      def clipWhenLowerLimitIsLessThanHigher(outputScaledValue, outputRange):
          if (outputScaledValue < outputRange[0]):
              return outputRange[0]
          elif (outputScaledValue > outputRange[1]):
              return outputRange[1]
          else:
              return outputScaledValue
          end
      end

      slope = computeSlope(rawRange, scaledRange)
      intercept = computeIntercept(slope, rawRange, scaledRange)
      scaledValue = slope * value + intercept
      return clipScaledValue(scaledValue, scaledRange)
  end

  def limit(value, range):
      return scale(value, range, range)
  end


  rq_init_comm_if_connected(9, "1")
  rq_init_comm_if_connected(2, "2")
  rq_init_comm_if_connected(3, "3")
  rq_init_comm_if_connected(4, "4")
  rq_print_connected_grippers()
  rq_gripper_communication_thread = run rq_gripper_communication()
  set_closed_norm(97.6470588235294, 1)
  set_open_norm(1.1764705882352942, 1)
  set_closed_mm(0.0, 1)
  set_open_mm(53.0, 1)
  set_closed_norm(100.0, 2)
  set_open_norm(0.0, 2)
  set_closed_mm(0.0, 2)
  set_open_mm(50.0, 2)
  set_closed_norm(100.0, 3)
  set_open_norm(0.0, 3)
  set_closed_mm(0.0, 3)
  set_open_mm(50.0, 3)
  set_closed_norm(100.0, 4)
  set_open_norm(0.0, 4)
  set_closed_mm(0.0, 4)
  set_open_mm(50.0, 4)
  rq_current_limit_enabled = False
  while(not rq_gripper_communication_thread_started):
      sync()
  end
  # end: URCap Installation Node
  # begin: URCap Installation Node
  #   Source: OPC UA, 2.0.2, Rocketfarm AS
  #   Type: OPC UA
  global opcua_daemon = rpc_factory("xmlrpc", "http://127.0.0.1:40409/RPC2")
  def opcua_client_connect(address):
  return opcua_daemon.client_connect(address)
  end
  def opcua_client_get_id(client_name):
  return opcua_daemon.client_get_id(client_name)
  end
  def opcua_client_try_connect(client_id):
  opcua_result = False
  if (opcua_daemon.client_connect(client_id)):
  sleep(0.01)
  opcua_result = opcua_daemon.client_is_connected(client_id)
  opcua_retry = 10
  while ( (not opcua_result) and (opcua_retry > 0) ):
  sleep(0.1)
  opcua_result = opcua_daemon.client_is_connected(client_id)
  opcua_retry = opcua_retry - 1
  end
  end
  return opcua_result
  end
  def opcua_client_disconnect(client_id):
  return opcua_daemon.client_disconnect(client_id)
  end
  def opcua_client_is_connected(client_id):
  return opcua_daemon.client_is_connected(client_id)
  end
  def opcua_client_read_byid(client_id, namespace_id, variable_id):
  return opcua_daemon.client_read_variable_by_id(client_id, namespace_id, variable_id)
  end
  def opcua_client_read_byname(client_id, namespace_id, variable_name):
  return opcua_daemon.client_read_variable_by_name(client_id, namespace_id, variable_name)
  end
  def opcua_client_write_byid(client_id, namespace_id, variable_id, variable_value):
  return opcua_daemon.client_write_variable_by_id(client_id, namespace_id, variable_id, variable_value)
  end
  def opcua_client_write_byname(client_id, namespace_id, variable_name, variable_value):
  return opcua_daemon.client_write_variable_by_name(client_id, namespace_id, variable_name, variable_value)
  end
  def opcua_client_last_error(client_id):
  return opcua_daemon.client_get_last_error(client_id)
  end
  def opcua_server_read_byname(variable_name):
  return opcua_daemon.server_read_variable_by_name(variable_name)
  end
  def opcua_server_write_byname(variable_name, variable_value):
  return opcua_daemon.server_write_variable_by_name(variable_name, variable_value)
  end
  def opcua_server_last_error():
  return opcua_daemon.server_get_last_error()
  end
  def opcua_error_to_string(errorCode):
  return opcua_daemon.error_code_to_string(errorCode)
  end
  # end: URCap Installation Node
  global CAM_Pose=p[0,0,0,0,0,0]
  global CAM_Relation=""
  global CMD_Abort=  False
  global CMD_Clear=  False
  global CMD_Reset=  False
  global CMD_Start=  False
  global CMD_Suspend=  False
  global CMD_Unhold=  False
  global CMD_Unsuspend=  False
  global CNT_Rack_Output=0
  global FNC_Freedrive=  False
  global PRC_TubCounter=0
  global STP=0
  global easyPickCount=0
  global easyPickCount_4=0
  global easyPickCount_6=0
  global easyPickCount_7=0
  global easyPickNoObj=0
  global easyPickNoObj_4=0
  global easyPickNoObj_6=0
  global easyPickNoObj_7=0
  global easyPickParts=0
  global easyPickParts_4=0
  global easyPickParts_6=0
  global easyPickParts_7=0
  global Container_mid_1_p=p[-.379239199143, -.127191311915, .299999999998, .000000000046, -.000000000021, -1.247199999994]
  global Container_mid_1_q=[-2.477408934449926, -1.2969853503591224, -1.875639182904262, -1.539621866126728, 1.5731943360401213, -2.8009955944022717]
  global Container_capt_p=p[-.525590029047, .407247642794, .411588185841, -.000000000107, .000000000065, -2.896148821900]
  global Container_capt_q=[-3.5968351615224767, -2.0050156108707204, -0.8176271154495112, -1.8895759482008394, 1.5730967555598792, -2.2743681102957645]
  global Waypoint_51_p=p[-.335468094724, -.217855817953, .299999999998, .000000000047, -.000000000014, -.994837065669]
  global Waypoint_51_q=[-2.2250460001249586, -1.2969853503591224, -1.875639182904262, -1.539621866126728, 1.573194336040121, -2.800995594402271]
  global Waypoint_13_p=p[-.479450777041, .284140798427, .125270103493, -.276792173670, 2.098433187455, -2.121256516887]
  global Waypoint_13_q=[-2.8915050665484827, -1.9549266300597132, -2.2318272590637207, -1.6654960117735804, 0.020810842514038086, -0.4019392172442835]
  global Waypoint_70_p=p[-.472820924464, .292439826304, .207418370234, -.259787347864, -2.053484648504, 2.070709755662]
  global Waypoint_70_q=[-2.969927421603815, -2.07168115810532, -1.6835546062719366, -2.4953958198513964, 0.4489790927922641, -0.005578998612037367]
  global Waypoint_2_p=p[-.312961047461, -.152991312519, .223609826854, -.745314530454, -1.713873240489, 1.673341715282]
  global Waypoint_2_q=[-2.3560472170459192, -2.183784624139303, -1.4583134651184082, -2.6435262165465296, 1.6522362232208252, 0.043451953679323196]
  global Waypoint_3_p=p[-.113749865836, -.390110151572, .317307487562, -.519383711706, -.839884211339, 1.756868173041]
  global Waypoint_3_q=[-1.8909733931170862, -1.720626016656393, -1.5115610361099243, -2.1240560017027796, 2.1809096336364746, 0.7227501273155212]
  global Waypoint_15_p=p[.029144035010, -.436802470887, .327885032028, -.521560953301, -.623641814548, 1.862659450154]
  global Waypoint_15_q=[-1.564817253743307, -1.556895188321807, -1.6826975345611572, -1.6944714985289515, 2.2362685203552246, 1.117417335510254]
  global Waypoint_14_p=p[.068712235638, -.569419545175, .285215357659, -.679242949116, -.712065334485, 1.394044574094]
  global Waypoint_14_q=[-1.5731792953485346, -1.8029235103747094, -1.6781008808776736, -1.2218450646111982, 2.4719572998240125, 1.6394218026856375]
  global Waypoint_4_p=p[-.047220457210, -.557624911767, .136370962514, -.679242949107, -.712065334475, 1.394044574096]
  global Waypoint_4_q=[-1.7740079055958748, -2.0023561428872334, -1.7577251142892676, -1.18903287716154, 2.4487287370345143, 1.322902469273079]
  global Waypoint_25_p=p[.065436479647, -.569388431626, .287820755049, -.679242949185, -.712065334557, 1.394044574070]
  global Waypoint_25_q=[-1.5789263550890595, -1.8020194754825436, -1.6702557537748035, -1.237882536889547, 2.471995808083492, 1.6301087487321393]
  global Waypoint_39_p=p[.137772150180, -.577759956854, .299999999946, .000000000217, -.000000000207, -1.594351842625]
  global Waypoint_39_q=[-1.108978697428574, -1.776486680444405, -1.413737665315093, -1.5218908901738937, 1.5733062372356947, -1.0863866394180182]
  global Waypoint_41_p=p[.074222967010, -.565641640647, .234620140366, -.516884386806, .529223682286, -1.529619060506]
  global Waypoint_41_q=[-0.9596722604286052, -1.8767069964135548, -1.4892746174057256, -1.7813862040292285, 1.0520698599867686, -0.8199687448260349]
  global Waypoint_40_p=p[.039987741677, -.564832865048, .191055405868, -.767560686167, .343136533060, -2.241315728308]
  global Waypoint_40_q=[-1.0070649180116558, -1.8745927522477324, -1.6139175023195245, -1.6337474788493545, 1.032708081143138, -0.11587278312988403]
  global Waypoint_42_p=p[.041363380882, -.564865360786, .192805844739, .278500165520, .624117100927, .762272396553]
  global Waypoint_42_q=[-1.0050718976263102, -1.8744386685524779, -1.609151451954446, -1.6399653140247947, 1.0334006002355505, -3.254032861659603]
  global Waypoint_43_p=p[.041363380886, -.564865360780, .192805844755, .854271020883, .226833028600, 2.453002871494]
  global Waypoint_43_q=[-1.0050567614299233, -1.874341297657562, -1.6092945416026048, -1.6397580431809713, 1.0333661149462194, -5.0371728933995605]
  global Waypoint_44_p=p[.040882892233, -.564854254876, .192193763716, .110913882012, .659173708659, .275719738520]
  global Waypoint_44_q=[-1.0057704811530535, -1.8745207681598055, -1.6107765025572558, -1.637858394640876, 1.033164860873599, -2.7487836132940755]
  global Waypoint_45_p=p[.042647731639, -.564895808997, .194439423694, -.451694728506, .563172064821, -1.343350300184]
  global Waypoint_45_q=[-1.0032860829914387, -1.8741561795270565, -1.6048483308761785, -1.6453689714776623, 1.0342050634514657, -1.06078829880322]
  global Waypoint_46_p=p[.099944144487, -.566244126804, .267342790130, -.451694834765, .563172023386, -1.343350532536]
  global Waypoint_46_q=[-0.9257438092434924, -1.889970530402497, -1.3828165217629076, -1.8916791100652528, 1.0664350961373816, -0.9805910833329659]
  global Waypoint_47_p=p[.099944144444, -.566244126727, .267342790273, -.101742139519, .058679218003, -1.457888523314]
  global Waypoint_47_q=[-1.1112623176383014, -1.729989471869196, -1.5530029871033957, -1.4442770617454777, 1.4670579052775654, -1.2224020460061675]
  global Waypoint_48_p=p[-.136182767566, -.647487115908, .294247768372, -.101742139549, .058679218020, -1.457888523312]
  global Waypoint_48_q=[-1.532196177857717, -1.9115932455375173, -1.2651848069729779, -1.5055651746702665, 1.4703193777418382, -1.646379689188814]
  global Waypoint_49_p=p[-.159024328559, -.641021381179, .047691706070, -.000000000033, -.000000000027, -1.457897102937]
  global Waypoint_49_q=[-1.6098490079965062, -2.1164987141784586, -1.6156631902166785, -0.9800092198841526, 1.573231151532669, -1.722204302767242]
  global Waypoint_50_p=p[-.159024328558, -.641021381151, .291114489351, -.000000000033, -.000000000027, -1.457897102937]
  global Waypoint_50_q=[-1.609190265995684, -1.9426985888940234, -1.2189094859258596, -1.55056435122874, 1.5734384912955113, -1.7235116759964022]
  global Waypoint_53_p=p[-.050111345339, -.357608435610, .335880801283, .034180375734, .020280946727, -.284888945062]
  global Waypoint_53_q=[-1.3262308189700454, -1.2221767968893875, -1.8246061249803773, -1.7046285947349489, 1.567288986353525, -2.612420684434543]
  global Spatula_above_p=p[.241880327671, -.243077591927, .290283157642, .000026293989, -.000477463062, 3.067686800856]
  global Spatula_above_q=[-0.3881264518731289, -1.1433094134493045, -1.996913957798169, -1.572030383936684, 1.5734346414190374, 1.2567789862982233]
  global Spatula_pick_p=p[.240292635430, -.243077591534, .189212061148, .000026293987, -.000477463065, 3.067686800855]
  global Spatula_pick_q=[-0.39083408330539005, -1.1777602778656497, -2.2383115866577645, -1.2961817529600745, 1.573403050820434, 1.2551372216266965]
  global container_start_p=p[.200650292946, -.570238751958, .366326773614, 1.360500828661, .021700128770, 2.681649891414]
  global container_start_q=[-0.7669977765142582, -2.188996679669204, -0.7412727239230232, -2.581362891432544, 1.0193601740278728, 1.1884911920528847]
  global container_wp_1_p=p[.170613637794, -.572150573676, .294509026043, 1.259497117139, -.008270589399, 2.787717865625]
  global container_wp_1_q=[-0.8129253370121727, -2.0726598902108755, -1.0846040680899218, -2.2403146195823957, 1.0281191187839607, 1.0435744211830564]
  global Waypoint_55_p=p[.077280900603, -.567308602990, .212067617714, 1.259497117148, -.008270589399, 2.787717865619]
  global Waypoint_55_q=[-0.9181858327853867, -1.9744793804952083, -1.4540279077890048, -1.9155621911627945, 0.9643238328181578, 0.9457250675800015]
  global Waypoint_56_p=p[.135568164031, -.570867938153, .245215470413, 1.476861317558, -.018269607491, 2.679642659499]
  global Waypoint_56_q=[-0.8259784040282607, -2.108036981522602, -1.2111990877342924, -2.2405969375728745, 0.9451797152137279, 1.125710531287379]
  global Waypoint_74_p=p[.164827890887, -.574638012411, .193751361296, 2.053636896063, -.046507887560, 2.274278266449]
  global Waypoint_74_q=[-0.7657213433975762, -2.450387120010788, -0.9886183070290357, -2.7078095590939375, 0.8831550681477878, 1.5106229631053527]
  global ftr_scoop2_p=p[.194287054614, -.495779761333, .282072128495, -.179029871953, 1.612108092436, -.016025695011]
  global ftr_scoop2_q=[-0.5957383150173561, -2.264100500923713, -1.1936887184643812, -2.8893702964346097, 0.8750688478879766, -1.4109843517598684]
  global aftr_scoo3_p=p[-.289759911340, -.315385007342, .303743796282, .159961590809, 1.627415489603, -.344855744095]
  global aftr_scoo3_q=[-1.3374747909924949, -1.6809733407851706, -1.9857606509106667, -2.713564895186775, 0.5589807453366573, -1.3631067603374376]
  global Waypoint_60_p=p[-.013316432876, -.544772031582, .383371643081, 2.208233379808, .037543335712, 2.097559881761]
  global Waypoint_60_q=[-0.9328326161883087, -2.0999933666355775, -1.1958015693111372, -3.060905141293654, 0.690378518537611, 1.7121940951337198]
  global Waypoint_61_p=p[-.412188693372, -.356446875193, .383371643081, 1.751740964455, -.739956256289, 1.600691174920]
  global Waypoint_61_q=[-1.766185342973321, -2.0999933666355775, -1.1958015693111372, -3.060905141293654, 0.690378518537611, 1.7121940951337198]
  global Waypoint_75_p=p[-.343126484123, -.342779621892, .335357223804, .359429517288, 1.600352990741, -.365083732359]
  global Waypoint_75_q=[-1.517806275013295, -1.8136828056045395, -1.737638081810795, -2.8432599585466436, 0.5149430839716123, -1.4579122147201877]
  global aftr_scoop1_p=p[.138503854266, -.514479969882, .214153672011, -.134825326227, 1.559916297527, -.059196589314]
  global aftr_scoop1_q=[-0.6880464314785328, -2.2689986529709643, -1.3310176475983653, -2.673087158390708, 0.8340516295138949, -1.4557846480003231]
  global After_disp_3_p=p[.125934854156, -.585611107804, .299545938076, .959554236104, -.134386766509, 2.880651774211]
  global After_disp_3_q=[-0.9434480594885066, -2.016473586333989, -1.1036579072158617, -2.096459283015281, 1.1479556364931514, 0.8433331387406042]
  global Waypoint_62_p=p[-.542658707241, -.114281911009, .251261544113, 1.813043609523, -.679411528034, 1.655271622964]
  global Waypoint_62_q=[-2.158300033470912, -1.9418836862428677, -1.8142999147147894, -2.778920736683023, 0.21900622104017292, 1.8983390235012934]
  global Waypoint_63_p=p[.101294795191, -.465376052375, .381756220355, .972633305146, -.158447626639, 2.887199602585]
  global Waypoint_63_q=[-0.8528172446194038, -1.7393709485118478, -1.2544079521837954, -2.2703112963960628, 1.1965892397133469, 0.91867216443391]
  global Start_p=p[-.033064633790, -.365398531763, .389873206922, .000000000001, .000000000001, 2.725785203584]
  global Start_q=[-1.287596562866887, -1.232866726886848, -1.6880113260231102, -1.7912103151657988, 1.5729028131945846, 0.6981423183093938]
  global Waypoint_76_p=p[-.479450777041, .284140798427, .125270103493, -.276792173670, 2.098433187454, -2.121256516887]
  global Waypoint_76_q=[-2.891505066548503, -1.9549266300590151, -2.231827259067863, -1.6654960117542226, 0.020810842514162875, -0.4019392172601952]
  global PowderA_wayp1_p=p[-.472820924474, .292439826233, .207418370237, -.137787250486, 2.177332259632, -2.152029714756]
  global PowderA_wayp1_q=[-2.911134078210732, -1.90240864358569, -1.968768330510411, -2.500365101593811, 0.11427687110891149, 0.0958980389250167]
  global Waypoint_80_p=p[-.303921889165, -.326082520111, .297721580072, -.584846481381, 1.914382606328, -1.960922301253]
  global Waypoint_80_q=[-1.6364180099980672, -2.041258366871811, -1.472153549517767, -2.7572808013122696, 0.9684003593854582, 0.047163023020230455]
  global Decapp_above_p=p[-.013480295948, -.359153355979, .266194408367, -.879653555922, 1.646336924805, -1.709111068605]
  global Decapp_above_q=[-0.9632157249872035, -2.0163405763031657, -1.5968194594157152, -2.6579215719847085, 1.251243398585566, 0.047906446502667066]
  global Decapp_place_p=p[-.013480295848, -.359153356116, .158558645017, -.879653554904, 1.646336919751, -1.709111066446]
  global Decapp_place_q=[-0.9633419174801583, -2.157735564881908, -1.695182597572722, -2.418253553201909, 1.2517436353048952, 0.04819090596102882]
  global Waypoint_78_p=p[-.051450028091, -.519555688329, .365718563414, -1.287302938145, 1.077637394477, -1.218524965834]
  global Waypoint_78_q=[-0.9214276262416012, -1.8899696965062578, -1.4939326452510562, -2.840015661555725, 0.5585157189668353, 0.033997638875617575]
  global Waypoint_81_p=p[-.030847790230, -.346237542439, .241203613248, .000000000000, .000000000000, .000000000000]
  global Waypoint_81_q=[-1.265848516232941, -1.1652881302267932, -2.11003646605462, -1.4369228603041853, 1.573284436504383, -2.835929896730388]
  global Waypoint_79_p=p[-.030847972829, -.346235312674, .229874122470, .000000000000, .000000000000, .000000000000]
  global Waypoint_79_q=[-1.2659333103898618, -1.1699230683425625, -2.1365870669440055, -1.4057372655396474, 1.5732787836040316, -2.8358953794066757]
  global Waypoint_82_p=p[-.031079593487, -.346547394534, .293012696855, -.000011575267, -.000017731224, -.000713984074]
  global Waypoint_82_q=[-1.2664169521879751, -1.1572597700415788, -1.982185304253158, -1.5727862504184884, 1.5732673022058234, -2.83632822711502]
  global Cap_above_p=p[-.163602500478, -.618357694237, .258271116068, .000026793591, -.000032305852, -.969382601663]
  global Cap_above_q=[-1.6181634639269902, -1.896432778341337, -1.3662765317923142, -1.449515114018281, 1.5734416863575176, -2.220489512402157]
  global Cap_Place_p=p[-.153420247224, -.637174247221, .035295616791, .000000000002, -.000000000002, -1.457849918374]
  global Cap_Place_q=[-1.6014084627078784, -2.123124488207292, -1.6429187572395012, -0.946127085055064, 1.573175527437006, -1.7136981844648291]
  global OP_PowderA2_p=p[.009371277507, -.409434369247, .294169017766, -.823281033205, 1.709410851243, -1.698303593897]
  global OP_PowderA2_q=[-0.9994544761745754, -2.1395254572673217, -1.3437567783153916, -2.8143375616690456, 1.2617899549595724, 0.019614613715634555]
  global OP_PowderA_abov_p=p[-.012145216791, -.363335041455, .315325728178, -.777135478411, 1.752984823781, -1.740925591659]
  global OP_PowderA_abov_q=[-1.01634425044037, -2.024785947780374, -1.4658894155189923, -2.8070189735738786, 1.3091674480404514, 0.020022086766872782]
  global OP_PowderA_pick_p=p[-.012145216707, -.363335041590, .179898787547, -.777135478413, 1.752984823781, -1.740925591659]
  global OP_PowderA_pick_q=[-1.0165129229305911, -2.176980100858497, -1.6127054339661555, -2.5080740815244567, 1.3098787614888208, 0.020270375244195882]
  global Op_PowA_wP_p=p[-.173727579245, -.372934016396, .295116627479, -.972390492433, 1.540962074418, -1.548745344994]
  global Op_PowA_wP_q=[-1.1740587397768483, -1.865656321049359, -1.7426943793777419, -2.679427276872525, 0.8588908769087338, 0.017944699631825187]
  global Waypoint_1_p=p[-.451048883256, -.340589460864, .308223661552, .097058877504, .091048998701, -1.578386010942]
  global Waypoint_1_q=[-2.222400490437643, -1.7554131946959437, -1.398173213005066, -1.6564461193480433, 1.5042352676391602, -2.2106884161578577]
  global Spatula_otw_p=p[-.038472058237, -.263141484147, .425351216717, -.000441582511, -.000128175490, 3.034387645854]
  global Spatula_otw_q=[-1.1888947506684495, -1.0083288774886814, -1.7052227056065874, -1.9984805067363443, 1.5730180972985317, 0.48793409320312264]
  global pick_spat_L_abv_p=p[.247376339171, -.151300871293, .298405979617, .000026293989, -.000477463062, 3.067686800856]
  global pick_spat_L_abv_q=[-0.07082187843937948, -0.9918336120099029, -2.048431407771396, -1.6719226065707566, 1.5735148227092874, 1.5739821706892307]
  global spat_L_pick_p=p[.244425006707, -.151048053384, .192288246285, .000026293989, -.000477463065, 3.067686800855]
  global spat_L_pick_q=[-0.07170850917614935, -0.9939169317558161, -2.3190151588645502, -1.3992549297298966, 1.573619586467819, 1.5742112847515592]
  global spat_L_lift_p=p[.247500241215, -.151291104039, .242146826477, .000026293989, -.000477463064, 3.067686800855]
  global spat_L_lift_q=[-0.07132168213116863, -0.9873531406871798, -2.1938095635783172, -1.531024644535787, 1.5736129628476565, 1.5740661231239859]
  global spat_L_side_p=p[.251772314117, -.093610100391, .242165935204, .000026293989, -.000477463064, 3.067686800855]
  global spat_L_side_q=[0.16311920731341095, -0.9159674867544636, -2.2202625845173465, -1.5759061264106862, 1.5736725172206427, 1.8084579794657634]
  global spat_L_up_p=p[.248631729748, -.094370561652, .425351216716, .000026293989, -.000477463065, 3.067686800855]
  global spat_L_up_q=[0.16435650344985986, -1.008385469590376, -1.7051729211515223, -1.9985780211252369, 1.5729805495343943, 1.8078858605162342]
  global spat_M_up_p=p[.246651483123, -.200758466677, .427983242435, .000026293988, -.000477463066, 3.067686800854]
  global spat_M_up_q=[-0.2488061154947081, -1.1388154682286178, -1.6405006043284098, -1.932909670500866, 1.5729930693357987, 1.394694958078517]
  global spat_M_pick_p=p[.243754824031, -.195909855689, .192274495860, .000026293989, -.000477463063, 3.067686800855]
  global spat_M_pick_q=[-0.2371047546337337, -1.0815273547611497, -2.2806002623741977, -1.3500947192370933, 1.573515135501001, 1.4088438823663394]
  global spat_S_up_p=p[.250500617207, -.246905508589, .391583682111, .000026293987, -.000477463068, 3.067686800854]
  global spat_S_up_q=[-0.3880360419879594, -1.1962881911765244, -1.7058643812256875, -1.8101014540154097, 1.5731545967396166, 1.2558061200976702]
  global spat_S_pick_p=p[.245173607467, -.244249950907, .193022226997, .000026293988, -.000477463064, 3.067686800854]
  global spat_S_pick_q=[-0.38836215799357987, -1.1880037605751017, -2.222350098157584, -1.30189927792612, 1.5733998957551099, 1.2575641527417636]
  def Sub_Vision_V18():
    $ 714 "Sub_Vision_V18" "noBreak"
    $ 715 "PreSettings"
    $ 716 "CAM_LM_Detected≔ False "
    global CAM_LM_Detected=  False
    $ 717 "CAM_Captures≔0"
    global CAM_Captures=0
    $ 718 "CAM_Pose≔p[0,0,0,0,0,0]"
    global CAM_Pose=p[0,0,0,0,0,0]
    $ 719 "CAM_LM_Refinmnt≔ False "
    global CAM_LM_Refinmnt=  False
    $ 720 "CAM_LM_Refined≔ False "
    global CAM_LM_Refined=  False
    $ 721 "CAM_LM_Deviatn≔p[0,0,0,0,0,0]"
    global CAM_LM_Deviatn=p[0,0,0,0,0,0]
    $ 722 "CAM_LM_ID≔0"
    global CAM_LM_ID=0
    $ 723 "CAM_Done≔ False "
    global CAM_Done=  False
    $ 724 "CAM_CNT_Obj≔0"
    global CAM_CNT_Obj=0
    $ 725 "CAM_Result = []"
    CAM_Result = []
    $ 726 "OBJ_Detected≔ False "
    global OBJ_Detected=  False
    $ 727 "FRM_Reference≔p[0,0,0,0,0,0]"
    global FRM_Reference=p[0,0,0,0,0,0]
    $ 728 "'=========='"
    # '=========='
    $ 729 "Switch Action"
    switch_1 = Action
    $ 730 "Case 13"
    if (13 == switch_1):
    elif (15 == switch_1):
      $ 848 "Case 15"
    elif (131 == switch_1):
      $ 894 "Case 131"
      $ 895 "Read (SensoPart)"
      $ 896 "Action_Info≔'search for landmark'"
      global Action_Info="search for landmark"
      $ 897 "CAM_LM≔CAM_LMs[4]"
      global CAM_LM=CAM_LMs[4]
      $ 898 "CAM_Relation≔CAM_LM.capture_relation"
      global CAM_Relation=CAM_LM.capture_relation
      $ 899 "go to capture pose"
      $ 902 "If ITM_ID≟1 and JIG≟7"
      if (ITM_ID == 1  and  JIG == 7):
        $ 903 "PSE_T≔uLM_Cap_SSRack"
        global PSE_T=uLM_Cap_SSRack
      else:
        $ 904 "ElseIf ITM_ID≟5 and JIG≟7"
        if (ITM_ID == 5  and  JIG == 7):
          $ 905 "PSE_T≔FRM_Cap_SSRack"
          global PSE_T=FRM_Cap_SSRack
        else:
          $ 906 "ElseIf ITM_ID≟13 and JIG≟7"
          if (ITM_ID == 13  and  JIG == 7):
            $ 907 "PSE_T≔FRM_pick_rack_const"
            global PSE_T=p[-0.5568395192387274,0.34423986364170267,0.44698620470146266,-1.0069110132199915E-6,3.378712467497258E-5,-8.002029546773325E-6]
          else:
            $ 908 "ElseIf ITM_ID≟1 and JIG≟15"
            if (ITM_ID == 1 and JIG == 15):
              $ 909 "MoveJ"
              $ 910 "Container_mid_1" "breakAfter"
              movej(get_inverse_kin(Container_mid_1_p, qnear=Container_mid_1_q), a=1.3962634015954636, v=1.0471975511965976, r=0.05)
              $ 911 "Container_capt" "breakAfter"
              movej(get_inverse_kin(Container_capt_p, qnear=Container_capt_q), a=1.3962634015954636, v=1.0471975511965976)
              $ 912 "PSE_T≔FRM_Container_S_const"
              global PSE_T=p[-0.510412665574981,0.40064363362973565,0.41159789496794374,-1.1370875604168537E-5,-3.643547521609506E-6,-2.896122366208473]
            else:
              $ 913 "ElseIf ITM_ID≟1 and JIG≟16"
              if (ITM_ID == 1  and  JIG == 16):
                $ 914 "MoveJ"
                $ 915 "Waypoint_51" "breakAfter"
                movej(get_inverse_kin(Waypoint_51_p, qnear=Waypoint_51_q), a=1.3962634015954636, v=1.0471975511965976, r=0.05)
                $ 917 "PSE_T≔FRM_Weigh_scale_const"
                global PSE_T=p[-0.3454891122972868,0.06305469656946562,0.547028193804949,1.63274868305228E-4,-7.686242288056818E-5,-2.2741025165393225]
              else:
                $ 918 "ElseIf ITM_ID≟1 and JIG≟17"
                if (ITM_ID == 1  and  JIG == 17):
                  $ 919 "MoveJ"
                  $ 920 "Waypoint_51" "breakAfter"
                  movej(get_inverse_kin(Waypoint_51_p, qnear=Waypoint_51_q), a=1.3962634015954636, v=1.0471975511965976, r=0.05)
                  $ 922 "PSE_T≔FRM_Weigh_scale_const"
                  global PSE_T=p[-0.3454891122972868,0.06305469656946562,0.547028193804949,1.63274868305228E-4,-7.686242288056818E-5,-2.2741025165393225]
                else:
                  $ 923 "ElseIf ITM_ID≟1 and JIG≟21"
                  if (ITM_ID == 1  and  JIG == 21):
                    $ 924 "MoveJ"
                    $ 925 "Waypoint_51" "breakAfter"
                    movej(get_inverse_kin(Waypoint_51_p, qnear=Waypoint_51_q), a=1.3962634015954636, v=1.0471975511965976, r=0.05)
                    $ 927 "PSE_T≔FRM_PoTS_const"
                    global PSE_T=p[-0.5211683440725288,-0.17068665293155189,0.5469908617304544,2.009713344566374E-4,5.545167142016751E-6,-2.2342044673695503]
                  end
                end
              end
            end
          end
        end
      end
      $ 928 "do_transition(PSE_T, keep_rxry=False)"
      do_transition(PSE_T, keep_rxry=False)
      $ 929 "Set"
      set_tcp(p[0.0,0.0,0.161,3.1415,0.0,0.0])
      $ 930 "MoveJ"
      $ 931 "PSE_T" "breakAfter"
      movej(PSE_T, a=1.3962634015954636, v=1.7453292519943295)
      $ 932 "CAM_Pose≔get_actual_tcp_pose()"
      global CAM_Pose= get_actual_tcp_pose ()
      $ 933 "Loop  not CAM_Done and  not ERROR.FLAG and  not CMD_Stop"
      while (  not  CAM_Done  and    not  ERROR.FLAG  and    not  CMD_Stop):
        $ 934 "adjust capture pose"
        $ 935 "If CAM_LM_Detected and CAM_LM_Refinmnt"
        if (CAM_LM_Detected  and  CAM_LM_Refinmnt):
          $ 936 "PSE_T≔p[0,0,0.300,0,0,0]"
          global PSE_T=p[0,0,0.300,0,0,0]
          $ 937 "CAM_Pose≔PSE_T"
          global CAM_Pose=PSE_T
          $ 938 "If  not is_reachable(FRM_Reference,[PSE_T])"
          if (  not  is_reachable(FRM_Reference,[PSE_T])):
            $ 939 "Error"
            $ 940 "set_error(ERROR_POSE_NOT_REACHABLE)"
            set_error(ERROR_POSE_NOT_REACHABLE)
          end
          $ 941 "If  not ERROR.FLAG"
          if (  not  ERROR.FLAG):
            $ 942 "MoveJ"
            $ 943 "PSE_T" "breakAfter"
            set_tcp(p[0.0,0.0,0.161,0.0,0.0,0.0])
            movej(pose_trans(FRM_Reference, PSE_T), a=0.8726646259971648, v=1.3962634015954636)
            $ 944 "CAM_LM_Refined≔ True "
            global CAM_LM_Refined=  True
          end
        else:
          $ 945 "ElseIf  not CAM_LM_Detected and CAM_Captures>0"
          if (  not  CAM_LM_Detected  and  CAM_Captures>0):
            $ 946 "MoveL"
            $ 947 "If FRM_Reference≟p[0,0,0,0,0,0]"
            if (FRM_Reference == p[0,0,0,0,0,0]):
              $ 948 "PSE_T≔get_random_pose(pose_ref=CAM_Pose, mode='cubic', range_max=[0.150,0.150,0.015])"
              global PSE_T=get_random_pose(pose_ref=CAM_Pose, mode="cubic", range_max=[0.150,0.150,0.015])
            else:
              $ 953 "Else" "noBreak"
              $ 954 "PSE_T≔get_random_pose(pose_ref=CAM_Pose, mode='rotation', range_max=[10,10,0])"
              global PSE_T=get_random_pose(pose_ref=CAM_Pose, mode="rotation", range_max=[10,10,0])
              $ 955 "CAM_LM_Refined≔ True "
              global CAM_LM_Refined=  True
            end
            $ 956 "If get_inverse_kin_has_solution(pose_trans(FRM_Reference, PSE_T))"
            if (get_inverse_kin_has_solution( pose_trans (FRM_Reference, PSE_T))):
              $ 957 "Comment"
              # Comment
              $ 958 "PSE_T" "breakAfter"
              set_tcp(p[0.0,0.0,0.161,3.1415,0.0,0.0])
              movel(pose_trans(FRM_Reference, PSE_T), a=0.03, v=0.05)
            else:
              $ 959 "Else" "noBreak"
              $ 960 "'If random pose is out of reach, set the initial cam pose'"
              # 'If random pose is out of reach, set the initial cam pose'
              $ 961 "PSE_T≔CAM_Pose"
              global PSE_T=CAM_Pose
            end
          end
        end
        $ 962 "Wait: 2.0"
        sleep(2.0)
        $ 963 "trigger"
        $ 964 "If ITM_ID≟1 and JIG≟7"
        if (ITM_ID == 1  and  JIG == 7):
          # begin: URCap Program Node
          #   Source: SensoPart VISOR Robotic, 2.0.0, SensoPart Industriesensorik GmbH
          #   Type: VISOR Trigger
          $ 965 "# 1 VISOR Trigger"
          visor_changeJob(1, "Landmark_INVITE_2", 6000)
          visor_trigger(1, 6000, "arm")
          # end: URCap Program Node
        else:
          $ 966 "ElseIf ITM_ID≟5 and JIG≟7"
          if (ITM_ID == 5  and  JIG == 7):
            # begin: URCap Program Node
            #   Source: SensoPart VISOR Robotic, 2.0.0, SensoPart Industriesensorik GmbH
            #   Type: VISOR Trigger
            $ 967 "# 1 VISOR Trigger"
            visor_changeJob(1, "Landmark_INVITE_2", 6000)
            visor_trigger(1, 6000, "arm")
            # end: URCap Program Node
          else:
            $ 968 "ElseIf ITM_ID≟13 and JIG≟7"
            if (ITM_ID == 13  and  JIG == 7):
              # begin: URCap Program Node
              #   Source: SensoPart VISOR Robotic, 2.0.0, SensoPart Industriesensorik GmbH
              #   Type: VISOR Trigger
              $ 969 "# 1 VISOR Trigger"
              visor_changeJob(1, "Landmark_INVITE_2", 6000)
              visor_trigger(1, 6000, "arm")
              # end: URCap Program Node
            else:
              $ 970 "ElseIf ITM_ID≟1 and JIG≟15"
              if (ITM_ID == 1 and JIG == 15):
                # begin: URCap Program Node
                #   Source: SensoPart VISOR Robotic, 2.0.0, SensoPart Industriesensorik GmbH
                #   Type: VISOR Trigger
                $ 971 "# 1 VISOR Trigger"
                visor_changeJob(1, "PowderA", 6000)
                visor_trigger(1, 6000, "arm")
                # end: URCap Program Node
              else:
                $ 972 "ElseIf ITM_ID≟1 and JIG≟16"
                if (ITM_ID == 1 and JIG == 16):
                  # begin: URCap Program Node
                  #   Source: SensoPart VISOR Robotic, 2.0.0, SensoPart Industriesensorik GmbH
                  #   Type: VISOR Trigger
                  $ 973 "# 1 VISOR Trigger"
                  visor_changeJob(1, "Weigh_target", 6000)
                  visor_trigger(1, 6000, "arm")
                  # end: URCap Program Node
                else:
                  $ 974 "ElseIf ITM_ID≟1 and JIG≟17"
                  if (ITM_ID == 1 and JIG == 17):
                    # begin: URCap Program Node
                    #   Source: SensoPart VISOR Robotic, 2.0.0, SensoPart Industriesensorik GmbH
                    #   Type: VISOR Trigger
                    $ 975 "# 1 VISOR Trigger"
                    visor_changeJob(1, "Weigh_target", 6000)
                    visor_trigger(1, 6000, "arm")
                    # end: URCap Program Node
                  else:
                    $ 976 "ElseIf ITM_ID≟1 and JIG≟21"
                    if (ITM_ID == 1 and JIG == 21):
                      # begin: URCap Program Node
                      #   Source: SensoPart VISOR Robotic, 2.0.0, SensoPart Industriesensorik GmbH
                      #   Type: VISOR Trigger
                      $ 977 "# 1 VISOR Trigger"
                      visor_changeJob(1, "Weigh_target", 6000)
                      visor_trigger(1, 6000, "arm")
                      # end: URCap Program Node
                    end
                  end
                end
              end
            end
          end
        end
        $ 981 "TM_3D_Found≔visor_partsFound(1)"
        global TM_3D_Found= visor_partsFound (1)
        $ 982 "If TM_3D_Found>0"
        if (TM_3D_Found>0):
          $ 983 "CAM_LM_Detected≔ True "
          global CAM_LM_Detected=  True
          $ 984 "CAM_Captures≔0"
          global CAM_Captures=0
        else:
          $ 985 "Else" "noBreak"
          $ 986 "CAM_LM_Detected≔ False "
          global CAM_LM_Detected=  False
          $ 987 "CAM_Captures≔CAM_Captures+1"
          global CAM_Captures=CAM_Captures+1
        end
        $ 992 "result"
        $ 993 "If CAM_LM_Detected"
        if (CAM_LM_Detected):
          $ 994 "If (CAM_LM_Refinmnt and CAM_LM_Refined) or  not CAM_LM_Refinmnt"
          if ((CAM_LM_Refinmnt  and  CAM_LM_Refined)  or    not  CAM_LM_Refinmnt):
            $ 1052 "If ITM_ID≟1 and JIG≟7"
            if (ITM_ID == 1  and  JIG == 7):
              $ 1053 "CAM_LM_SSRack≔visor_getPose3d(1, 0)"
              global CAM_LM_SSRack= visor_getPose3d (1, 0)
            else:
              $ 1054 "ElseIf ITM_ID≟5 and JIG≟7"
              if (ITM_ID == 5  and  JIG == 7):
                $ 1055 "CAM_LM_SSRack≔visor_getPose3d(1, 0)"
                global CAM_LM_SSRack= visor_getPose3d (1, 0)
              else:
                $ 1056 "ElseIf ITM_ID≟13 and JIG≟7"
                if (ITM_ID == 13  and  JIG == 7):
                  $ 1057 "CAM_LM_Bott≔visor_getPose3d(1, 0)"
                  global CAM_LM_Bott= visor_getPose3d (1, 0)
                else:
                  $ 1058 "ElseIf ITM_ID≟1 and JIG≟15"
                  if (ITM_ID == 1 and JIG == 15):
                    $ 1059 "CAM_LM_Cont_S≔visor_getPose3d(1, 0)"
                    global CAM_LM_Cont_S= visor_getPose3d (1, 0)
                    $ 1060 "cont_img_pose≔get_actual_tcp_pose()"
                    global cont_img_pose= get_actual_tcp_pose ()
                  else:
                    $ 1061 "ElseIf ITM_ID≟1 and JIG≟16"
                    if (ITM_ID == 1 and JIG == 16):
                      $ 1062 "CAM_cont≔visor_getPose3d(1, 0)"
                      global CAM_cont= visor_getPose3d (1, 0)
                      $ 1063 "cont_img_pose≔get_actual_tcp_pose()"
                      global cont_img_pose= get_actual_tcp_pose ()
                    else:
                      $ 1064 "ElseIf ITM_ID≟1 and JIG≟17"
                      if (ITM_ID == 1 and JIG == 17):
                        $ 1066 "cont_img_pose≔get_actual_tcp_pose()"
                        global cont_img_pose= get_actual_tcp_pose ()
                      else:
                        $ 1067 "ElseIf ITM_ID≟1 and JIG≟21"
                        if (ITM_ID == 1 and JIG == 21):
                          $ 1069 "cont_img_pose≔get_actual_tcp_pose()"
                          global cont_img_pose= get_actual_tcp_pose ()
                        end
                      end
                    end
                  end
                end
              end
            end
            $ 1070 "CAM_Done≔ True "
            global CAM_Done=  True
          end
        else:
          $ 1071 "ElseIf  not CAM_LM_Detected and CAM_Captures<CAM_PRM_Retries"
          if (  not  CAM_LM_Detected  and  CAM_Captures<CAM_PRM_Retries):
            $ 1072 "CAM_LM_Refined≔ False "
            global CAM_LM_Refined=  False
          else:
            $ 1073 "ElseIf CAM_Captures≥CAM_PRM_Retries"
            if (CAM_Captures >= CAM_PRM_Retries):
              $ 1074 "CAM_Done≔ True "
              global CAM_Done=  True
              $ 1075 "Error"
              $ 1076 "set_error(ERROR_NO_LANDMARK)"
              set_error(ERROR_NO_LANDMARK)
            end
          end
        end
      end
    elif (151 == switch_1):
      $ 1077 "Case 151"
      $ 1078 "Detect (SensoPart)"
      $ 1079 "go to capture pose"
      $ 1080 "FRM_Reference≔FRM_Cap_SSRack"
      global FRM_Reference=FRM_Cap_SSRack
      $ 1081 "PSE_T≔p[0,0,-0.00,0,0,0]"
      global PSE_T=p[0,0,-0.00,0,0,0]
      $ 1082 "do_transition(pose_trans(FRM_Reference, PSE_T), keep_rxry=False)"
      do_transition( pose_trans (FRM_Reference, PSE_T), keep_rxry=False)
      $ 1083 "JNT_Q≔get_actual_joint_positions()"
      global JNT_Q= get_actual_joint_positions ()
      $ 1084 "JNT_Q≔[JNT_Q[0], JNT_Q[1], JNT_Q[2], JNT_Q[3], JNT_Q[4], 0]"
      global JNT_Q=[JNT_Q[0], JNT_Q[1], JNT_Q[2], JNT_Q[3], JNT_Q[4], 0]
      $ 1085 "Set"
      set_tcp(p[0.0,0.0,0.161,3.1415,0.0,0.0])
      $ 1086 "movej(get_inverse_kin(pose_trans(FRM_Reference, PSE_T), qnear=JNT_Q))"
      movej(get_inverse_kin( pose_trans (FRM_Reference, PSE_T), qnear=JNT_Q))
      $ 1087 "CAM_Pose≔pose_trans(pose_inv(FRM_Reference), get_actual_tcp_pose())"
      global CAM_Pose= pose_trans ( pose_inv (FRM_Reference),  get_actual_tcp_pose ())
      $ 1088 "Loop  not CAM_Done and  not ERROR.FLAG and  not CMD_Stop"
      while (  not  CAM_Done  and    not  ERROR.FLAG  and    not  CMD_Stop):
        $ 1089 "If  not OBJ_Detected and CAM_Captures>0"
        if (  not  OBJ_Detected  and  CAM_Captures>0):
          $ 1090 "MoveL"
          $ 1091 "If FRM_Reference≟p[0,0,0,0,0,0]"
          if (FRM_Reference == p[0,0,0,0,0,0]):
            $ 1093 "PSE_T≔get_random_pose(pose_ref=CAM_Pose, mode='rotation', range_max=[15,15,0])"
            global PSE_T=get_random_pose(pose_ref=CAM_Pose, mode="rotation", range_max=[15,15,0])
          else:
            $ 1094 "Else" "noBreak"
            $ 1095 "PSE_T≔get_random_pose(pose_ref=CAM_Pose, mode='rotation', range_max=[10,10,0])"
            global PSE_T=get_random_pose(pose_ref=CAM_Pose, mode="rotation", range_max=[10,10,0])
          end
          $ 1096 "If get_inverse_kin_has_solution(pose_trans(FRM_Reference, PSE_T))"
          if (get_inverse_kin_has_solution( pose_trans (FRM_Reference, PSE_T))):
            $ 1097 "PSE_T" "breakAfter"
            set_tcp(p[0.0,0.0,0.161,3.1415,0.0,0.0])
            movel(pose_trans(FRM_Reference, PSE_T), a=0.03, v=0.05)
          else:
            $ 1098 "Else" "noBreak"
            $ 1099 "'If random pose is out of reach, set the initial cam pose'"
            # 'If random pose is out of reach, set the initial cam pose'
            $ 1100 "PSE_T≔CAM_Pose"
            global PSE_T=CAM_Pose
            $ 1101 "PSE_T" "breakAfter"
            set_tcp(p[0.0,0.0,0.161,3.1415,0.0,0.0])
            movel(pose_trans(FRM_Reference, PSE_T), a=0.03, v=0.05)
          end
        end
        $ 1102 "Wait: 0.5"
        sleep(0.5)
        $ 1103 "Set"
        set_tcp(p[0.0,0.0,0.161,3.1415,0.0,0.0])
        # begin: URCap Program Node
        #   Source: SensoPart VISOR Robotic, 2.0.0, SensoPart Industriesensorik GmbH
        #   Type: VISOR Trigger
        $ 1104 "# 1 VISOR Trigger"
        visor_changeJob(1, "Object Detection Single", 6000)
        visor_trigger(1, 6000, "arm")
        # end: URCap Program Node
        $ 1105 "If visor_isResponseOk(1)"
        if ( visor_isResponseOk (1)):
          $ 1106 "CAM_CNT_Obj≔visor_partsFound(1)"
          global CAM_CNT_Obj= visor_partsFound (1)
          $ 1107 "CAM_OBJ_Pose≔visor_getPose3d(1, 0)"
          global CAM_OBJ_Pose= visor_getPose3d (1, 0)
          $ 1108 "If CAM_CNT_Obj>0"
          if (CAM_CNT_Obj>0):
            $ 1109 "CAM_OBJ_Color≔visor_getAdditionalData(1, 0)"
            global CAM_OBJ_Color= visor_getAdditionalData (1, 0)
            $ 1110 "CAM_DetectScore≔to_num(visor_getAdditionalData(1, 1))/1000"
            global CAM_DetectScore=to_num( visor_getAdditionalData (1, 1))/1000
            $ 1111 "OBJ_Detected≔ True "
            global OBJ_Detected=  True
          end
        else:
          $ 1112 "Else" "noBreak"
          $ 1113 "CAM_Captures≔CAM_Captures+1"
          global CAM_Captures=CAM_Captures+1
        end
        $ 1114 "If OBJ_Detected"
        if (OBJ_Detected):
          $ 1115 "Get object data"
          $ 1116 "PRC_CntDetect≔0"
          global PRC_CntDetect=0
          $ 1117 "Loop PRC_CntDetect<CAM_CNT_Obj"
          while (PRC_CntDetect<CAM_CNT_Obj):
            $ 1118 "get object and jig number"
            $ 1119 "If ITM_ID≟1 and JIG≟7"
            if (ITM_ID == 1  and  JIG == 7):
              $ 1120 "FRM_Reference≔FRM_Cap_SSRack"
              global FRM_Reference=FRM_Cap_SSRack
            else:
              $ 1121 "ElseIf ITM_ID≟5 and JIG≟7"
              if (ITM_ID == 5  and  JIG == 7):
                $ 1122 "FRM_Reference≔uLM_Cap_SSRack"
                global FRM_Reference=uLM_Cap_SSRack
              end
            end
            $ 1125 "PSE_T≔pose_trans(pose_inv(FRM_Reference), CAM_OBJ_Pose)"
            global PSE_T= pose_trans ( pose_inv (FRM_Reference), CAM_OBJ_Pose)
            $ 1126 "CAM_Result.append(get_pattern_counter(PSE_T, 'X', pattern=[10, 5], patternsize=[0.181, 0.081]))"
            CAM_Result.append(get_pattern_counter(PSE_T, "X", pattern=[10, 5], patternsize=[0.181, 0.081]))
            $ 1127 "PRC_CntDetect≔PRC_CntDetect+1"
            global PRC_CntDetect=PRC_CntDetect+1
          end
          $ 1128 "CAM_Done≔ True "
          global CAM_Done=  True
        else:
          $ 1129 "ElseIf CAM_Captures≥CAM_PRM_Retries"
          if (CAM_Captures >= CAM_PRM_Retries):
            $ 1130 "CAM_Done≔ True "
            global CAM_Done=  True
          else:
            $ 1131 "Else" "noBreak"
            $ 1132 "CAM_Captures≔CAM_Captures+1"
            global CAM_Captures=CAM_Captures+1
          end
        end
      end
    end
    $ 1133 "'=========='"
    # '=========='
    $ 1134 "PostSettings"
    $ 1135 "FRM_Reference≔p[0,0,0,0,0,0]"
    global FRM_Reference=p[0,0,0,0,0,0]
    $ 1136 "Set"
    set_tcp(p[0.0,0.0,0.161,3.1415,0.0,0.0])
    $ 1137 "CAM_Pose≔p[0,0,0,0,0,0]"
    global CAM_Pose=p[0,0,0,0,0,0]
    $ 1138 "Action≔0"
    global Action=0
    $ 1139 "Action_Info≔''"
    global Action_Info=""
  end
  def Sub_Action_V4():
    $ 1140 "Sub_Action_V4" "noBreak"
    $ 1141 "PreSettings"
    $ 1142 "init poses"
    $ 1143 "PSE_A≔p[0,0,0,0,0,0]"
    global PSE_A=p[0,0,0,0,0,0]
    $ 1144 "PSE_A_H≔p[0,0,0,0,0,0]"
    global PSE_A_H=p[0,0,0,0,0,0]
    $ 1145 "PSE_T≔p[0,0,0,0,0,0]"
    global PSE_T=p[0,0,0,0,0,0]
    $ 1146 "PSE_T_H≔p[0,0,0,0,0,0]"
    global PSE_T_H=p[0,0,0,0,0,0]
    $ 1147 "PSE_G≔p[0,0,0,0,0,0]"
    global PSE_G=p[0,0,0,0,0,0]
    $ 1148 "PSE_G_H≔p[0,0,0,0,0,0]"
    global PSE_G_H=p[0,0,0,0,0,0]
    $ 1149 "PSE_R≔p[0,0,0,0,0,0]"
    global PSE_R=p[0,0,0,0,0,0]
    $ 1150 "PSE_R_H≔p[0,0,0,0,0,0]"
    global PSE_R_H=p[0,0,0,0,0,0]
    $ 1151 "JNT_Q≔[0,0,0,0,0,0]"
    global JNT_Q=[0,0,0,0,0,0]
    $ 1152 "JNT_S≔[0,0,0,0,0,0]"
    global JNT_S=[0,0,0,0,0,0]
    $ 1153 "Gripping parameters"
    $ 1154 "OBJ = find_object_by_type(OBJs, OBJ_Type)"
    OBJ = find_object_by_type(OBJs, OBJ_Type)
    $ 1155 "GRP_Open_Pos≔OBJ.dimension.diameter * 1000 + 6"
    global GRP_Open_Pos=OBJ.dimension.diameter * 1000 + 6
    $ 1156 "GRP_Offset≔OBJ.gripper_offset"
    global GRP_Offset=OBJ.gripper_offset
    $ 1157 "rq_set_force_norm(50)"
     rq_set_force_norm (50)
    $ 1158 "rq_set_speed_norm(50)"
     rq_set_speed_norm (50)
    $ 1159 "Switch ITM_ID"
    switch_1 = ITM_ID
    $ 1160 "Case 1"
    if (1 == switch_1):
      $ 1161 "uML"
      $ 1162 "JIG2 = find_object_by_type(JIGs, JIG)"
      JIG2 = find_object_by_type(JIGs, JIG)
      $ 1163 "JIG_Offset≔JIG2.jig_offset"
      global JIG_Offset=JIG2.jig_offset
      $ 1164 "Switch JIG"
      switch_2 = JIG
      $ 1165 "Case 1"
      if (1 == switch_2):
        $ 1166 "3FG"
        $ 1167 "define poses"
        $ 1168 "FRM_Reference≔ULM_3FG"
        global FRM_Reference=ULM_3FG
        $ 1169 "JNT_Q≔JNT_HOME"
        global JNT_Q=JNT_HOME
        $ 1170 "PSE_T≔pose_trans(GRP_Offset, JIG_Offset)"
        global PSE_T= pose_trans (GRP_Offset, JIG_Offset)
        $ 1171 "PSE_A≔pose_trans(PSE_T, p[0,0,0.100,0,0,0])"
        global PSE_A= pose_trans (PSE_T, p[0,0,0.100,0,0,0])
        $ 1172 "PSE_R≔pose_add(PSE_T, p[0,0,0.100,0,0,0])"
        global PSE_R= pose_add (PSE_T, p[0,0,0.100,0,0,0])
      elif (2 == switch_2):
        $ 1173 "Case 2"
        $ 1174 "Input"
        $ 1175 "'CHANGE THE REFERENCE TO THE FRAME TO MOVE IN'"
        # 'CHANGE THE REFERENCE TO THE FRAME TO MOVE IN'
        $ 1176 "define poses"
        $ 1177 "FRM_Reference≔ULM_Input"
        global FRM_Reference=ULM_Input
        $ 1178 "PSE_T≔pose_trans(pose_trans(get_pattern_pos_rectangle(OBJ_Nbr, 'X', [10,5], patternsize=[0.181,0.081]), GRP_Offset), JIG_Offset)"
        global PSE_T= pose_trans ( pose_trans (get_pattern_pos_rectangle(OBJ_Nbr, "X", [10,5], patternsize=[0.181,0.081]), GRP_Offset), JIG_Offset)
        $ 1179 "If Action≟1"
        if (Action == 1):
          $ 1180 "PSE_R≔pose_add(PSE_T, p[0,0,0.200,0,0,0])"
          global PSE_R= pose_add (PSE_T, p[0,0,0.200,0,0,0])
          $ 1181 "PSE_A≔pose_add(PSE_T, p[0,0,0.100,0,0,0])"
          global PSE_A= pose_add (PSE_T, p[0,0,0.100,0,0,0])
        else:
          $ 1182 "ElseIf Action≟2"
          if (Action == 2):
            $ 1183 "PSE_R≔pose_add(PSE_T, p[0,0,0.100,0,0,0])"
            global PSE_R= pose_add (PSE_T, p[0,0,0.100,0,0,0])
            $ 1184 "PSE_A≔pose_add(PSE_T, p[0,0,0.200,0,0,0])"
            global PSE_A= pose_add (PSE_T, p[0,0,0.200,0,0,0])
          end
        end
      elif (3 == switch_2):
        $ 1185 "Case 3"
        $ 1186 "Output"
        $ 1187 "'CHANGE THE REFERENCE TO THE FRAME TO MOVE IN'"
        # 'CHANGE THE REFERENCE TO THE FRAME TO MOVE IN'
        $ 1188 "define poses"
        $ 1189 "FRM_Reference≔ULM_Output"
        global FRM_Reference=ULM_Output
        $ 1190 "PSE_T≔pose_trans(pose_trans(get_pattern_pos_rectangle(OBJ_Nbr, 'X', [10,5], patternsize=[0.181,0.081]), GRP_Offset), JIG_Offset)"
        global PSE_T= pose_trans ( pose_trans (get_pattern_pos_rectangle(OBJ_Nbr, "X", [10,5], patternsize=[0.181,0.081]), GRP_Offset), JIG_Offset)
        $ 1192 "If Action≟1"
        if (Action == 1):
          $ 1193 "PSE_R≔pose_add(PSE_T, p[0,0,0.200,0,0,0])"
          global PSE_R= pose_add (PSE_T, p[0,0,0.200,0,0,0])
          $ 1194 "PSE_A≔pose_add(PSE_T, p[0,0,0.100,0,0,0])"
          global PSE_A= pose_add (PSE_T, p[0,0,0.100,0,0,0])
        else:
          $ 1195 "ElseIf Action≟2"
          if (Action == 2):
            $ 1196 "PSE_R≔pose_add(PSE_T, p[0,0,0.100,0,0,0])"
            global PSE_R= pose_add (PSE_T, p[0,0,0.100,0,0,0])
            $ 1197 "PSE_A≔pose_add(PSE_T, p[0,0,0.200,0,0,0])"
            global PSE_A= pose_add (PSE_T, p[0,0,0.200,0,0,0])
          end
        end
      elif (4 == switch_2):
        $ 1198 "Case 4"
        $ 1199 "jig centrifuge racks"
        $ 1200 "define poses"
        $ 1201 "FRM_Reference≔ULM_Cent_Racks"
        global FRM_Reference=ULM_Cent_Racks
        $ 1202 "PSE_T≔get_pattern_pos_rectangle(JIG_Slot, 'X', [4,1], patternsize=[0.291,0])"
        global PSE_T=get_pattern_pos_rectangle(JIG_Slot, "X", [4,1], patternsize=[0.291,0])
        $ 1203 "If OBJ_Nbr≠0"
        if (OBJ_Nbr != 0):
          $ 1204 "PSE_T≔pose_trans(pose_trans(PSE_T, get_pattern_pos_rectangle(OBJ_Nbr, 'X', [3,3], patternsize=[0.060,0.060])),p[-0.030, -0.030,0,0,0,3.927])"
          global PSE_T= pose_trans ( pose_trans (PSE_T, get_pattern_pos_rectangle(OBJ_Nbr, "X", [3,3], patternsize=[0.060,0.060])),p[-0.030, -0.030,0,0,0,3.927])
        end
        $ 1205 "PSE_T≔pose_trans(PSE_T, GRP_Offset)"
        global PSE_T= pose_trans (PSE_T, GRP_Offset)
        $ 1206 "If Action≟1"
        if (Action == 1):
          $ 1207 "PSE_R≔pose_add(PSE_T, p[0,0,0.200,0,0,0])"
          global PSE_R= pose_add (PSE_T, p[0,0,0.200,0,0,0])
          $ 1208 "PSE_A≔pose_add(PSE_T, p[0,0,0.100,0,0,0])"
          global PSE_A= pose_add (PSE_T, p[0,0,0.100,0,0,0])
        else:
          $ 1209 "ElseIf Action≟2"
          if (Action == 2):
            $ 1210 "PSE_R≔pose_add(PSE_T, p[0,0,0.100,0,0,0])"
            global PSE_R= pose_add (PSE_T, p[0,0,0.100,0,0,0])
            $ 1211 "PSE_A≔pose_add(PSE_T, p[0,0,0.200,0,0,0])"
            global PSE_A= pose_add (PSE_T, p[0,0,0.200,0,0,0])
          end
        end
      elif (6 == switch_2):
        $ 1212 "Case 6"
        $ 1213 "Caps bin"
        $ 1214 "define poses"
        $ 1215 "'Drop cap'"
        # 'Drop cap'
        $ 1216 "FRM_Reference=ULM_Cap_Bin"
        FRM_Reference=ULM_Cap_Bin
        $ 1217 "PSE_T≔pose_RPY2RotVec(p[0,0,0,0,0,0])"
        global PSE_T=pose_RPY2RotVec(p[0,0,0,0,0,0])
        $ 1218 "PSE_T_H≔pose_add(PSE_T, p[0,0,-0.011,0,0,0])"
        global PSE_T_H= pose_add (PSE_T, p[0,0,-0.011,0,0,0])
        $ 1219 "PSE_A≔pose_trans(PSE_T, p[0,0,0.1,0,0,0])"
        global PSE_A= pose_trans (PSE_T, p[0,0,0.1,0,0,0])
        $ 1220 "PSE_R_H≔pose_add(PSE_T, p[0,0,0.100,0,0,0])"
        global PSE_R_H= pose_add (PSE_T, p[0,0,0.100,0,0,0])
        $ 1221 "PSE_R≔pose_add(PSE_T, p[0,0,0.100,0,0,0])"
        global PSE_R= pose_add (PSE_T, p[0,0,0.100,0,0,0])
      elif (7 == switch_2):
        $ 1222 "Case 7"
        $ 1223 "Sarstedt"
        $ 1224 "'CHANGE THE REFERENCE TO THE FRAME TO MOVE IN'"
        # 'CHANGE THE REFERENCE TO THE FRAME TO MOVE IN'
        $ 1230 "If TASK.ID≟10"
        if (TASK.ID == 10):
          $ 1231 "Frame & Position Params"
          $ 1233 "FRM_Reference = CAM_LM_SSRack"
          FRM_Reference = CAM_LM_SSRack
          $ 1238 "PSE_T≔uLM_SS_PickPlc"
          global PSE_T=uLM_SS_PickPlc
          $ 1239 "PSE_A≔pose_trans(PSE_T, p[0,0,0.1,0,0,0])"
          global PSE_A= pose_trans (PSE_T, p[0,0,0.1,0,0,0])
          $ 1240 "PSE_R≔pose_add(PSE_T, p[0,0,0.1,0,0,0])"
          global PSE_R= pose_add (PSE_T, p[0,0,0.1,0,0,0])
        else:
          $ 1241 "ElseIf TASK.ID≟11"
          if (TASK.ID == 11):
            $ 1242 "FRM_Reference = ULM_SS_Jig"
            FRM_Reference = ULM_SS_Jig
            $ 1243 "PSE_T≔pose_RPY2RotVec(p[0,0,0,0,0,0])"
            global PSE_T=pose_RPY2RotVec(p[0,0,0,0,0,0])
            $ 1244 "PSE_T≔pose_trans(PSE_T, GRP_Offset)"
            global PSE_T=pose_trans(PSE_T, GRP_Offset)
            $ 1245 "PSE_A≔pose_trans(PSE_T, p[0,0,0.1,0,0,0])"
            global PSE_A= pose_trans (PSE_T, p[0,0,0.1,0,0,0])
            $ 1246 "PSE_R≔pose_add(PSE_T, p[0,0,0.2,0,0,0])"
            global PSE_R= pose_add (PSE_T, p[0,0,0.2,0,0,0])
          end
        end
      elif (8 == switch_2):
        $ 1247 "Case 8"
        $ 1248 "NoK"
        $ 1249 "define poses"
        $ 1250 "'NoK'"
        # 'NoK'
        $ 1251 "FRM_Reference=ULM_NoK"
        FRM_Reference=ULM_NoK
        $ 1252 "PSE_T≔pose_RPY2RotVec(p[0,0,0,0,0,0])"
        global PSE_T=pose_RPY2RotVec(p[0,0,0,0,0,0])
        $ 1253 "PSE_A≔pose_trans(PSE_T, p[0,0,0.1,0,0,0])"
        global PSE_A= pose_trans (PSE_T, p[0,0,0.1,0,0,0])
        $ 1254 "PSE_R≔pose_add(PSE_T, p[0,0,0.100,0,0,0])"
        global PSE_R= pose_add (PSE_T, p[0,0,0.100,0,0,0])
      elif (9 == switch_2):
        $ 1255 "Case 9"
        $ 1256 "Pick_bott_jig"
        $ 1257 "define poses"
        $ 1258 "'NoK'"
        # 'NoK'
        $ 1259 "FRM_Reference=ULM_bottle_pick_const"
        FRM_Reference=p[0.08175869478771049,-0.47602162643540935,0.09,0.00141829700319658,-0.0027789445191063835,0.07763675748118615]
        $ 1260 "PSE_T≔pose_RPY2RotVec(p[0,0,0,0,0,0])"
        global PSE_T=pose_RPY2RotVec(p[0,0,0,0,0,0])
        $ 1261 "PSE_A≔pose_trans(PSE_T, p[0,0,0.1,0,0,0])"
        global PSE_A= pose_trans (PSE_T, p[0,0,0.1,0,0,0])
        $ 1262 "PSE_R≔pose_add(PSE_T, p[0,0,0.100,0,0,0])"
        global PSE_R= pose_add (PSE_T, p[0,0,0.100,0,0,0])
      elif (10 == switch_2):
        $ 1263 "Case 10"
        $ 1264 "Place_bott_jig"
        $ 1265 "define poses"
        $ 1266 "'NoK'"
        # 'NoK'
        $ 1267 "FRM_Reference=ULM_bottle_plac_const"
        FRM_Reference=p[-0.09502738395762109,-0.5154087721098056,0.095,0.0014590126708889871,-0.0028280855286173575,0.07763149296298452]
        $ 1268 "PSE_T≔pose_RPY2RotVec(p[0,0,0,0,0,0])"
        global PSE_T=pose_RPY2RotVec(p[0,0,0,0,0,0])
        $ 1269 "PSE_A≔pose_trans(PSE_T, p[0,0,0.1,0,0,0])"
        global PSE_A= pose_trans (PSE_T, p[0,0,0.1,0,0,0])
        $ 1270 "PSE_R≔pose_add(PSE_T, p[0,0,0.100,0,0,0])"
        global PSE_R= pose_add (PSE_T, p[0,0,0.100,0,0,0])
      elif (11 == switch_2):
        $ 1271 "Case 11"
        $ 1272 "Place_bott_jig"
        $ 1273 "define poses"
        $ 1274 "'NoK'"
        # 'NoK'
        $ 1275 "FRM_Reference=shake"
        FRM_Reference=shake
        $ 1276 "PSE_T≔pose_RPY2RotVec(p[0,0,0,0,0,0])"
        global PSE_T=pose_RPY2RotVec(p[0,0,0,0,0,0])
        $ 1277 "PSE_A≔pose_trans(PSE_T, p[0,0,0,0,0,0])"
        global PSE_A= pose_trans (PSE_T, p[0,0,0,0,0,0])
        $ 1278 "PSE_R≔pose_add(PSE_T, p[0,0,0,0,0,0])"
        global PSE_R= pose_add (PSE_T, p[0,0,0,0,0,0])
      elif (12 == switch_2):
        $ 1279 "Case 12"
        $ 1280 "Pick_Vial_jig"
        $ 1281 "define poses"
        $ 1282 "'NoK'"
        # 'NoK'
        $ 1283 "FRM_Reference=shake"
        FRM_Reference=shake
        $ 1284 "PSE_T≔pose_RPY2RotVec(p[0,0,0,0,0,0])"
        global PSE_T=pose_RPY2RotVec(p[0,0,0,0,0,0])
        $ 1285 "PSE_A≔pose_trans(PSE_T, p[0,0,0,0,0,0])"
        global PSE_A= pose_trans (PSE_T, p[0,0,0,0,0,0])
        $ 1286 "PSE_R≔pose_add(PSE_T, p[0,0,0,0,0,0])"
        global PSE_R= pose_add (PSE_T, p[0,0,0,0,0,0])
      end
    elif (2 == switch_1):
      $ 1287 "Case 2"
      $ 1288 "Centrifuge"
      $ 1289 "'CHANGE THE REFERENCE TO THE FRAME TO MOVE IN'"
      # 'CHANGE THE REFERENCE TO THE FRAME TO MOVE IN'
      $ 1290 "define poses"
      $ 1291 "FRM_Reference≔FRM_Centrifuge"
      global FRM_Reference=FRM_Centrifuge
      $ 1292 "PSE_T≔GRP_Offset"
      global PSE_T=GRP_Offset
      $ 1293 "If Action≟8"
      if (Action == 8):
        $ 1294 "PSE_R≔pose_add(PSE_T, p[0,0,0.250,0,0,0])"
        global PSE_R= pose_add (PSE_T, p[0,0,0.250,0,0,0])
        $ 1295 "PSE_A≔pose_add(PSE_T, p[0,0,0.150,0,0,0])"
        global PSE_A= pose_add (PSE_T, p[0,0,0.150,0,0,0])
      else:
        $ 1296 "ElseIf Action≟7"
        if (Action == 7):
          $ 1297 "PSE_R≔pose_add(PSE_T, p[0,0,0.150,0,0,0])"
          global PSE_R= pose_add (PSE_T, p[0,0,0.150,0,0,0])
          $ 1298 "PSE_A≔pose_add(PSE_T, p[0,0,0.250,0,0,0])"
          global PSE_A= pose_add (PSE_T, p[0,0,0.250,0,0,0])
        end
      end
    elif (3 == switch_1):
      $ 1299 "Case 3"
      $ 1300 "Output"
      $ 1301 "'CHANGE THE REFERENCE TO THE FRAME TO MOVE IN'"
      # 'CHANGE THE REFERENCE TO THE FRAME TO MOVE IN'
      $ 1302 "define poses"
      $ 1303 "FRM_Reference≔Base_const"
      global FRM_Reference=p[0.0,0.0,0.0,0.0,0.0,0.0]
      $ 1304 "PSE_T≔p[0,0,0,0,0,0]"
      global PSE_T=p[0,0,0,0,0,0]
      $ 1305 "PSE_A≔pose_add(PSE_T, p[0,0,0.150,0,0,0])"
      global PSE_A= pose_add (PSE_T, p[0,0,0.150,0,0,0])
      $ 1306 "PSE_R≔pose_add(PSE_T, p[0,0,0.100,0,0,0])"
      global PSE_R= pose_add (PSE_T, p[0,0,0.100,0,0,0])
    elif (5 == switch_1):
      $ 1307 "Case 5"
      $ 1308 "Sarstedt Pickup Table"
      $ 1309 "'CHANGE THE REFERENCE TO THE FRAME TO MOVE IN'"
      # 'CHANGE THE REFERENCE TO THE FRAME TO MOVE IN'
      $ 1310 "Switch JIG"
      switch_2 = JIG
      $ 1311 "Case 7"
      if (7 == switch_2):
        $ 1324 "Sarstedt"
        $ 1325 "'CHANGE THE REFERENCE TO THE FRAME TO MOVE IN'"
        # 'CHANGE THE REFERENCE TO THE FRAME TO MOVE IN'
        $ 1331 "If TASK.ID≟10"
        if (TASK.ID == 10):
          $ 1332 "Frame & Position Params"
          $ 1333 "FRM_Reference = CAM_LM_SSRack"
          FRM_Reference = CAM_LM_SSRack
          $ 1334 "PSE_T≔uLM_SS_PickPlc"
          global PSE_T=uLM_SS_PickPlc
          $ 1335 "PSE_A≔pose_trans(PSE_T, p[0,0,0.1,0,0,0])"
          global PSE_A= pose_trans (PSE_T, p[0,0,0.1,0,0,0])
          $ 1336 "PSE_R≔pose_add(PSE_T, p[0,0,0.1,0,0,0])"
          global PSE_R= pose_add (PSE_T, p[0,0,0.1,0,0,0])
        end
      end
    elif (13 == switch_1):
      $ 1343 "Case 13"
      $ 1344 "Sarstedt Pickup Table"
      $ 1345 "'CHANGE THE REFERENCE TO THE FRAME TO MOVE IN'"
      # 'CHANGE THE REFERENCE TO THE FRAME TO MOVE IN'
      $ 1346 "Switch JIG"
      switch_2 = JIG
      $ 1347 "Case 7"
      if (7 == switch_2):
        $ 1360 "Bottle"
        $ 1361 "'CHANGE THE REFERENCE TO THE FRAME TO MOVE IN'"
        # 'CHANGE THE REFERENCE TO THE FRAME TO MOVE IN'
        $ 1367 "If TASK.ID≟43"
        if (TASK.ID == 43):
          $ 1368 "Frame & Position Params"
          $ 1369 "FRM_Reference = CAM_LM_Bott"
          FRM_Reference = CAM_LM_Bott
          $ 1370 "PSE_T≔uLM_SS_PickPlc"
          global PSE_T=uLM_SS_PickPlc
          $ 1371 "PSE_A≔pose_trans(PSE_T, p[0,0,0.1,0,0,0])"
          global PSE_A= pose_trans (PSE_T, p[0,0,0.1,0,0,0])
          $ 1372 "PSE_R≔pose_add(PSE_T, p[0,0,0.1,0,0,0])"
          global PSE_R= pose_add (PSE_T, p[0,0,0.1,0,0,0])
        end
      end
    end
    $ 1379 "Additional check"
    $ 1380 "If  not is_reachable(FRM_Reference,[PSE_A,PSE_A_H,PSE_T,PSE_T_H,PSE_R,PSE_R_H])"
    if (  not  is_reachable(FRM_Reference,[PSE_A,PSE_A_H,PSE_T,PSE_T_H,PSE_R,PSE_R_H])):
      $ 1381 "Error"
      $ 1382 "set_error(ERROR_POSE_NOT_REACHABLE)"
      set_error(ERROR_POSE_NOT_REACHABLE)
      $ 1383 "Action≔0"
      global Action=0
    end
    $ 1384 "'=========='"
    # '=========='
    $ 1385 "Switch Action"
    switch_1 = Action
    $ 1386 "Case 1"
    if (1 == switch_1):
      $ 1387 "Pick"
      $ 1388 "Action_Info≔'pick object'"
      global Action_Info="pick object"
      $ 1389 "do_transition(pose_trans(FRM_Reference, PSE_T), keep_rxry=OBJ_Picked)"
      do_transition( pose_trans (FRM_Reference, PSE_T), keep_rxry=OBJ_Picked)
      $ 1390 "EOAT"
      $ 1391 "If  not OBJ_Picked"
      if (  not  OBJ_Picked):
        $ 1392 "rq_move_and_wait_mm(GRP_Open_Pos)"
         rq_move_and_wait_mm (GRP_Open_Pos)
      end
      $ 1393 "If PSE_A_H≠PSE_Z"
      if (PSE_A_H != PSE_Z):
        $ 1394 "If JNT_Q≠JNT_Z"
        if (JNT_Q != JNT_Z):
          $ 1395 "movej(get_inverse_kin(pose_trans(FRM_Reference, PSE_A_H), qnear=JNT_Q), r=0.050)"
          movej(get_inverse_kin( pose_trans (FRM_Reference, PSE_A_H), qnear=JNT_Q), r=0.050)
        else:
          $ 1396 "Else" "noBreak"
          $ 1397 "movej(pose_trans(FRM_Reference, PSE_A_H), r=0.050)"
          movej( pose_trans (FRM_Reference, PSE_A_H), r=0.050)
        end
      end
      $ 1398 "If PSE_A≠PSE_Z"
      if (PSE_A != PSE_Z):
        $ 1399 "If JNT_Q≠JNT_Z"
        if (JNT_Q != JNT_Z):
          $ 1400 "movej(get_inverse_kin(pose_trans(FRM_Reference, PSE_A), qnear=JNT_Q), r=0.020)"
          movej(get_inverse_kin( pose_trans (FRM_Reference, PSE_A), qnear=JNT_Q), r=0.020)
        else:
          $ 1401 "Else" "noBreak"
          $ 1402 "movej(pose_trans(FRM_Reference, PSE_A), r=0.020)"
          movej( pose_trans (FRM_Reference, PSE_A), r=0.020)
        end
      end
      $ 1403 "MoveL"
      $ 1404 "If PSE_T_H≠PSE_Z"
      if (PSE_T_H != PSE_Z):
        $ 1405 "PSE_T_H" "breakAfter"
        movel(pose_trans(FRM_Reference, PSE_T_H), a=0.5, v=0.4, r=0.01)
      end
      $ 1406 "PSE_T" "breakAfter"
      movel(pose_trans(FRM_Reference, PSE_T), a=0.08, v=0.12)
      $ 1407 "EOAT"
      $ 1408 "rq_set_force_norm(50)"
       rq_set_force_norm (50)
      $ 1409 "rq_close_and_wait()"
       rq_close_and_wait ()
      $ 1410 "OBJ_Picked≔rq_is_object_detected()"
      global OBJ_Picked= rq_is_object_detected ()
      $ 1411 "If  not OBJ_Picked"
      if (  not  OBJ_Picked):
        $ 1412 "set_error(ERROR_NO_OBJECT_TO_PICK)"
        set_error(ERROR_NO_OBJECT_TO_PICK)
      end
      $ 1413 "EXTT"
      $ 1414 "Switch JIG"
      switch_2 = JIG
      $ 1415 "Case 1"
      if (1 == switch_2):
        $ 1416 "3FG"
        $ 1417 "If OBJ_Picked"
        if (OBJ_Picked):
          $ 1418 "Set GRP_3F_Open=On"
          set_standard_digital_out(5, True)
        end
      end
      $ 1419 "If PSE_R_H≠PSE_Z"
      if (PSE_R_H != PSE_Z):
        $ 1420 "PSE_R" "breakAfter"
        movel(pose_trans(FRM_Reference, PSE_R), a=0.5, v=0.4, r=0.01)
        $ 1421 "PSE_R_H" "breakAfter"
        movel(pose_trans(FRM_Reference, PSE_R_H), a=0.5, v=0.4)
      else:
        $ 1422 "Else" "noBreak"
        $ 1423 "PSE_R" "breakAfter"
        movel(pose_trans(FRM_Reference, PSE_R), a=0.5, v=0.4)
      end
    elif (2 == switch_1):
      $ 1424 "Case 2"
    elif (3 == switch_1):
      $ 1466 "Case 3"
    elif (4 == switch_1):
      $ 1469 "Case 4"
    elif (6 == switch_1):
      $ 1472 "Case 6"
    elif (7 == switch_1):
      $ 1487 "Case 7"
    elif (8 == switch_1):
      $ 1516 "Case 8"
    elif (11 == switch_1):
      $ 1549 "Case 11"
    elif (12 == switch_1):
      $ 1586 "Case 12"
    elif (15 == switch_1):
      $ 1637 "Case 15"
    elif (30 == switch_1):
      $ 1640 "Case 30"
    elif (31 == switch_1):
      $ 1673 "Case 31"
    elif (32 == switch_1):
      $ 1685 "Case 32"
    elif (33 == switch_1):
      $ 1726 "Case 33"
    elif (35 == switch_1):
      $ 1792 "Case 35"
      $ 1793 "Pick the powder container"
      # begin: URCap Program Node
      #   Source: SensoPart VISOR Robotic, 2.0.0, SensoPart Industriesensorik GmbH
      #   Type: VISOR Robotic App
      $ 1796 "VISOR Easy Pick"
      def visorFuncEasyPick_a89ad0():
        # begin: URCap Program Node
        #   Source: SensoPart VISOR Robotic, 2.0.0, SensoPart Industriesensorik GmbH
        #   Type: Easy Pick Setup
        $ 1797 "# 1 Setup" "noBreak"
        local easyPickVisorId = 1
        local easyPickArmMounted = True
        local easyPickSetJob = True
        local easyPickJobName = "Container"
        local easyPickAtImgAcq = False
        local easyPickImgAcqPose = cont_img_pose
        # end: URCap Program Node
        # begin: URCap Program Node
        #   Source: SensoPart VISOR Robotic, 2.0.0, SensoPart Industriesensorik GmbH
        #   Type: Process
        $ 1798 "Process" "noBreak"
        local easyPickObjTaken = False
        local easyPickTrigger = False
        local easyPickPoseIdx = 0
        local easyPickPose = p[0,0,0,0,0,0]
        def easyPickFuncTrigger(visorId, setJob, jobName, arm):
        if (setJob):
          visor_changeJob(visorId, jobName, 6000)
        end
        if (arm):
          visor_trigger(visorId, 6000, "arm")
        else:
          visor_trigger(visorId, 6000)
        end
        global easyPickParts=visor_partsFound(visorId)
        visor_easyPickUpdate(visorId, "parts", visor_partsFound(visorId))
        return visor_getPose3d(visorId, 0)
      end
      while (not easyPickObjTaken):
        easyPickTrigger = (easyPickCount >= visor_partsFound(easyPickVisorId)) or (easyPickCount > 9) or (not visor_easyPickCheckIdent("6318e7", easyPickVisorId))
        if (easyPickTrigger):
          easyPickCount = 0
        end
        easyPickPoseIdx = easyPickCount
        easyPickPose = visor_getPose3d(easyPickVisorId, easyPickPoseIdx)
        visor_easyPickUpdate(easyPickVisorId, "counter", easyPickPoseIdx)
        # begin: URCap Program Node
        #   Source: SensoPart VISOR Robotic, 2.0.0, SensoPart Industriesensorik GmbH
        #   Type: Image Acquisition Pose
        $ 1799 "Image Acquisition Pose" "noBreak"
        if (easyPickTrigger):
          if (not easyPickAtImgAcq):
            movej(pose_trans(easyPickImgAcqPose,p[0.0000,0.0000,-0.0000,0.0000,0.0000,0.0000]),a=1.3963,v=1.0472,t=0.000000,r=0.000000)
            easyPickAtImgAcq = True
          end
          easyPickPose = easyPickFuncTrigger(easyPickVisorId, easyPickSetJob, easyPickJobName, easyPickArmMounted)
        end
        # end: URCap Program Node
        # begin: URCap Program Node
        #   Source: SensoPart VISOR Robotic, 2.0.0, SensoPart Industriesensorik GmbH
        #   Type: Object Detected
        $ 1800 "Object Detected" "noBreak"
        if (visor_partsFound(easyPickVisorId) > 0):
          $ 1801 "Open Gripper" "noBreak"
          # begin: URCap Program Node
          #   Source: Robotiq_Grippers, 1.8.4.4844, Robotiq Inc.
          #   Type: Gripper
          $ 1802 "Gripper Open (1)" "noBreak"
          if not(gripper_connected[0]):
            popup("Gripper 1 must be connected to run this program.", "No connection", False, True, True)
          end
          if not(rq_is_gripper_activated("1")):
            popup("Gripper 1 is not activated. Go to Installation tab > Gripper to activate it and run the program again.", "Not activated", False, True, True)
          end
          rq_set_pos_spd_for(0, 102, 77, "1")
          rq_wait_pos_spe_for_request(0, 102, 77, "1")
          rq_go_to("1")
          rq_wait("1")
          # end: URCap Program Node
          $ 1803 "MoveJ" "noBreak"
          $ 1804 "Waypoint_13" "noBreak"
          movej(get_inverse_kin(Waypoint_13_p, qnear=Waypoint_13_q), a=1.3962634015954636, v=1.0471975511965976)
          # begin: URCap Program Node
          #   Source: SensoPart VISOR Robotic, 2.0.0, SensoPart Industriesensorik GmbH
          #   Type: Approach Pose
          $ 1805 "Approach Pose" "noBreak"
          movej(pose_trans(easyPickPose,p[0.0000,0.0000,0.0500,0.0000,0.0000,0.0000]),a=1.3963,v=1.0472,t=0.000000,r=0.000000)
          # end: URCap Program Node
          # begin: URCap Program Node
          #   Source: SensoPart VISOR Robotic, 2.0.0, SensoPart Industriesensorik GmbH
          #   Type: Target Pose
          $ 1806 "Target Pose" "noBreak"
          movel(pose_trans(easyPickPose,p[0.0000,0.0000,-0.0000,0.0000,0.0000,0.0000]),a=0.5000,v=0.2500,t=0.000000,r=0.000000)
          # end: URCap Program Node
          $ 1807 "Close Gripper" "noBreak"
          # begin: URCap Program Node
          #   Source: Robotiq_Grippers, 1.8.4.4844, Robotiq Inc.
          #   Type: Gripper
          $ 1808 "Gripper Close (1)" "noBreak"
          if not(gripper_connected[0]):
            popup("Gripper 1 must be connected to run this program.", "No connection", False, True, True)
          end
          if not(rq_is_gripper_activated("1")):
            popup("Gripper 1 is not activated. Go to Installation tab > Gripper to activate it and run the program again.", "Not activated", False, True, True)
          end
          rq_set_pos_spd_for(255, 102, 77, "1")
          rq_wait_pos_spe_for_request(255, 102, 77, "1")
          rq_go_to("1")
          rq_wait("1")
          # end: URCap Program Node
          # begin: URCap Program Node
          #   Source: SensoPart VISOR Robotic, 2.0.0, SensoPart Industriesensorik GmbH
          #   Type: Exit Pose
          $ 1809 "Exit Pose" "noBreak"
          movel(pose_trans(easyPickPose,p[0.0000,0.0000,0.0500,0.0000,0.0000,0.0000]),a=0.5000,v=0.2500,t=0.000000,r=0.000000)
          # end: URCap Program Node
          easyPickObjTaken = True
        end
        # end: URCap Program Node
        # begin: URCap Program Node
        #   Source: SensoPart VISOR Robotic, 2.0.0, SensoPart Industriesensorik GmbH
        #   Type: No Object Detected
        $ 1810 "No Object Detected" "noBreak"
        if (visor_partsFound(easyPickVisorId) < 1):
          $ 1811 "Popup: No Container detected" "noBreak"
          popup("No Container detected", "Message", False, False, blocking=True)
          else:
        end
        # end: URCap Program Node
      end
      easyPickCount = easyPickCount + 1
      visor_easyPickUpdate(easyPickVisorId, "counter", easyPickCount)
      visor_easyPickSetIdent("6318e7", easyPickVisorId)
      # end: URCap Program Node
    end
    visorFuncEasyPick_a89ad0()
    # end: URCap Program Node
    $ 1812 "MoveJ"
    $ 1814 "Waypoint_70" "breakAfter"
    movej(get_inverse_kin(Waypoint_70_p, qnear=Waypoint_70_q), a=0.6981317007977318, v=0.5235987755982988)
    $ 1815 "Waypoint_2" "breakAfter"
    movej(get_inverse_kin(Waypoint_2_p, qnear=Waypoint_2_q), a=0.8726646259971648, v=0.5235987755982988, r=0.05)
    $ 1816 "Waypoint_3" "breakAfter"
    movej(get_inverse_kin(Waypoint_3_p, qnear=Waypoint_3_q), a=0.6981317007977318, v=0.5235987755982988, r=0.05)
    $ 1817 "MoveL"
    $ 1818 "Waypoint_15" "breakAfter"
    movel(Waypoint_15_p, a=0.5, v=0.1, r=0.05)
    $ 1819 "Waypoint_14" "breakAfter"
    movel(Waypoint_14_p, a=0.3, v=0.1)
    $ 1820 "Waypoint_4" "breakAfter"
    movel(Waypoint_4_p, a=0.3, v=0.05)
    # begin: URCap Program Node
    #   Source: Robotiq_Grippers, 1.8.4.4844, Robotiq Inc.
    #   Type: Gripper
    $ 1821 "Gripper Open (1)"
    if not(gripper_connected[0]):
      popup("Gripper 1 must be connected to run this program.", "No connection", False, True, True)
    end
    if not(rq_is_gripper_activated("1")):
      popup("Gripper 1 is not activated. Go to Installation tab > Gripper to activate it and run the program again.", "Not activated", False, True, True)
    end
    rq_set_pos_spd_for(0, 102, 77, "1")
    rq_wait_pos_spe_for_request(0, 102, 77, "1")
    rq_go_to("1")
    rq_wait("1")
    # end: URCap Program Node
    $ 1822 "MoveL"
    $ 1823 "Waypoint_25" "breakAfter"
    movel(Waypoint_25_p, a=0.3, v=0.1)
    $ 1824 "Waypoint_15" "breakAfter"
    movel(Waypoint_15_p, a=0.5, v=0.1, r=0.05)
    $ 1825 "Home (Safe)"
    movej([-1.2302089344500047, -1.2969853503591224, -1.875639182904262, -1.539621866126728, 1.5731943360401213, -2.80099559440227], a=1.3962634015954636, v=1.0471975511965976)
  elif (36 == switch_1):
    $ 1855 "Case 36"
    $ 1859 "Decap"
    $ 1897 "MoveJ"
    $ 1898 "Waypoint_39" "breakAfter"
    movej(get_inverse_kin(Waypoint_39_p, qnear=Waypoint_39_q), a=1.3962634015954636, v=1.0471975511965976)
    $ 1899 "MoveL"
    $ 1900 "Waypoint_41" "breakAfter"
    movel(Waypoint_41_p, a=0.5, v=0.1)
    $ 1901 "Waypoint_40" "breakAfter"
    movel(Waypoint_40_p, a=0.3, v=0.05)
    # begin: URCap Program Node
    #   Source: Robotiq_Grippers, 1.8.4.4844, Robotiq Inc.
    #   Type: Gripper
    $ 1902 "Gripper Close (1)"
    if not(gripper_connected[0]):
      popup("Gripper 1 must be connected to run this program.", "No connection", False, True, True)
    end
    if not(rq_is_gripper_activated("1")):
      popup("Gripper 1 is not activated. Go to Installation tab > Gripper to activate it and run the program again.", "Not activated", False, True, True)
    end
    rq_set_pos_spd_for(255, 77, 51, "1")
    rq_wait_pos_spe_for_request(255, 77, 51, "1")
    rq_go_to("1")
    rq_wait("1")
    # end: URCap Program Node
    $ 1903 "Loop 2 times"
    Loop_2 = 0
    while (Loop_2 < 2):
      $ 1904 "MoveL"
      $ 1905 "Waypoint_42" "breakAfter"
      movel(Waypoint_42_p, a=1.2, v=0.5)
      $ 1906 "Waypoint_43" "breakAfter"
      movel(Waypoint_43_p, a=1.2, v=0.25)
      # begin: URCap Program Node
      #   Source: Robotiq_Grippers, 1.8.4.4844, Robotiq Inc.
      #   Type: Gripper
      $ 1907 "Gripper Move40mm (1)"
      if not(gripper_connected[0]):
        popup("Gripper 1 must be connected to run this program.", "No connection", False, True, True)
      end
      if not(rq_is_gripper_activated("1")):
        popup("Gripper 1 is not activated. Go to Installation tab > Gripper to activate it and run the program again.", "Not activated", False, True, True)
      end
      rq_set_pos_spd_for(63, 77, 51, "1")
      rq_wait_pos_spe_for_request(63, 77, 51, "1")
      rq_go_to("1")
      rq_wait("1")
      # end: URCap Program Node
      $ 1908 "MoveL"
      $ 1909 "Waypoint_44" "breakAfter"
      movel(Waypoint_44_p, a=1.2, v=0.5)
      $ 1910 "Waypoint_45" "breakAfter"
      movel(Waypoint_45_p, a=1.2, v=0.25)
      # begin: URCap Program Node
      #   Source: Robotiq_Grippers, 1.8.4.4844, Robotiq Inc.
      #   Type: Gripper
      $ 1911 "Gripper Move11mm (1)"
      if not(gripper_connected[0]):
        popup("Gripper 1 must be connected to run this program.", "No connection", False, True, True)
      end
      if not(rq_is_gripper_activated("1")):
        popup("Gripper 1 is not activated. Go to Installation tab > Gripper to activate it and run the program again.", "Not activated", False, True, True)
      end
      rq_set_pos_spd_for(200, 77, 51, "1")
      rq_wait_pos_spe_for_request(200, 77, 51, "1")
      rq_go_to("1")
      rq_wait("1")
      # end: URCap Program Node
      Loop_2 = Loop_2 + 1
    end
    $ 1912 "MoveL"
    $ 1913 "Waypoint_46" "breakAfter"
    movel(Waypoint_46_p, a=0.3, v=0.05)
    $ 1914 "Waypoint_47" "breakAfter"
    movel(Waypoint_47_p, a=0.5, v=0.1)
    $ 1915 "Waypoint_48" "breakAfter"
    movel(Waypoint_48_p, a=1.2, v=0.25)
    $ 1916 "Waypoint_49" "breakAfter"
    movel(Waypoint_49_p, a=1.2, v=0.25)
    # begin: URCap Program Node
    #   Source: Robotiq_Grippers, 1.8.4.4844, Robotiq Inc.
    #   Type: Gripper
    $ 1917 "Gripper Move35mm (1)"
    if not(gripper_connected[0]):
      popup("Gripper 1 must be connected to run this program.", "No connection", False, True, True)
    end
    if not(rq_is_gripper_activated("1")):
      popup("Gripper 1 is not activated. Go to Installation tab > Gripper to activate it and run the program again.", "Not activated", False, True, True)
    end
    rq_set_pos_spd_for(87, 77, 51, "1")
    rq_wait_pos_spe_for_request(87, 77, 51, "1")
    rq_go_to("1")
    rq_wait("1")
    # end: URCap Program Node
    $ 1918 "MoveL"
    $ 1919 "Waypoint_50" "breakAfter"
    movel(Waypoint_50_p, a=1.2, v=0.25)
    $ 1920 "Home (Safe)"
    movej([-1.2302089344500047, -1.2969853503591224, -1.875639182904262, -1.539621866126728, 1.5731943360401213, -2.80099559440227], a=1.3962634015954636, v=1.0471975511965976)
  elif (37 == switch_1):
    $ 1921 "Case 37"
    $ 1922 "Powder dispensing"
    $ 1923 "zero_scale()"
    zero_scale()
    # begin: URCap Program Node
    #   Source: SensoPart VISOR Robotic, 2.0.0, SensoPart Industriesensorik GmbH
    #   Type: VISOR Robotic App
    $ 1924 "VISOR Easy Pick"
    def visorFuncEasyPick_5fe5fa():
      # begin: URCap Program Node
      #   Source: SensoPart VISOR Robotic, 2.0.0, SensoPart Industriesensorik GmbH
      #   Type: Easy Pick Setup
      $ 1925 "# 1 Setup" "noBreak"
      local easyPickVisorId = 1
      local easyPickArmMounted = True
      local easyPickSetJob = True
      local easyPickJobName = "Weigh_scale"
      local easyPickAtImgAcq = False
      local easyPickImgAcqPose = cont_img_pose
      # end: URCap Program Node
      # begin: URCap Program Node
      #   Source: SensoPart VISOR Robotic, 2.0.0, SensoPart Industriesensorik GmbH
      #   Type: Process
      $ 1926 "Process" "noBreak"
      local easyPickObjTaken = False
      local easyPickTrigger = False
      local easyPickPoseIdx = 0
      local easyPickPose = p[0,0,0,0,0,0]
      def easyPickFuncTrigger(visorId, setJob, jobName, arm):
      if (setJob):
        visor_changeJob(visorId, jobName, 6000)
      end
      if (arm):
        visor_trigger(visorId, 6000, "arm")
      else:
        visor_trigger(visorId, 6000)
      end
      global easyPickParts_4=visor_partsFound(visorId)
      visor_easyPickUpdate(visorId, "parts", visor_partsFound(visorId))
      return visor_getPose3d(visorId, 0)
    end
    while (not easyPickObjTaken):
      easyPickTrigger = (easyPickCount_4 >= visor_partsFound(easyPickVisorId)) or (easyPickCount_4 > 9) or (not visor_easyPickCheckIdent("a3cf6b", easyPickVisorId))
      if (easyPickTrigger):
        easyPickCount_4 = 0
      end
      easyPickPoseIdx = easyPickCount_4
      easyPickPose = visor_getPose3d(easyPickVisorId, easyPickPoseIdx)
      visor_easyPickUpdate(easyPickVisorId, "counter", easyPickPoseIdx)
      # begin: URCap Program Node
      #   Source: SensoPart VISOR Robotic, 2.0.0, SensoPart Industriesensorik GmbH
      #   Type: Image Acquisition Pose
      $ 1927 "Image Acquisition Pose" "noBreak"
      if (easyPickTrigger):
        if (not easyPickAtImgAcq):
          movej(pose_trans(easyPickImgAcqPose,p[0.0000,0.0000,-0.0000,0.0000,0.0000,0.0000]),a=1.3963,v=1.0472,t=0.000000,r=0.000000)
          easyPickAtImgAcq = True
        end
        easyPickPose = easyPickFuncTrigger(easyPickVisorId, easyPickSetJob, easyPickJobName, easyPickArmMounted)
      end
      # end: URCap Program Node
      # begin: URCap Program Node
      #   Source: SensoPart VISOR Robotic, 2.0.0, SensoPart Industriesensorik GmbH
      #   Type: Object Detected
      $ 1928 "Object Detected" "noBreak"
      if (visor_partsFound(easyPickVisorId) > 0):
        $ 1929 "Open Gripper" "noBreak"
        $ 1930 "MoveL" "noBreak"
        $ 1931 "Weight_value≔get_weight()" "noBreak"
        global Weight_value=get_weight()
        # begin: URCap Program Node
        #   Source: Robotiq_Grippers, 1.8.4.4844, Robotiq Inc.
        #   Type: Gripper
        $ 1932 "Gripper Open (1)" "noBreak"
        if not(gripper_connected[0]):
          popup("Gripper 1 must be connected to run this program.", "No connection", False, True, True)
        end
        if not(rq_is_gripper_activated("1")):
          popup("Gripper 1 is not activated. Go to Installation tab > Gripper to activate it and run the program again.", "Not activated", False, True, True)
        end
        rq_set_pos_spd_for(0, 77, 77, "1")
        rq_wait_pos_spe_for_request(0, 77, 77, "1")
        rq_go_to("1")
        rq_wait("1")
        # end: URCap Program Node
        $ 1933 "Waypoint_53" "noBreak"
        movel(Waypoint_53_p, a=0.6, v=0.15, r=0.05)
        $ 1934 "Spatula_above" "noBreak"
        movel(Spatula_above_p, a=0.6, v=0.15)
        $ 1935 "Spatula_pick" "noBreak"
        movel(Spatula_pick_p, a=0.6, v=0.15)
        # begin: URCap Program Node
        #   Source: Robotiq_Grippers, 1.8.4.4844, Robotiq Inc.
        #   Type: Gripper
        $ 1936 "Gripper Close (1)" "noBreak"
        if not(gripper_connected[0]):
          popup("Gripper 1 must be connected to run this program.", "No connection", False, True, True)
        end
        if not(rq_is_gripper_activated("1")):
          popup("Gripper 1 is not activated. Go to Installation tab > Gripper to activate it and run the program again.", "Not activated", False, True, True)
        end
        rq_set_pos_spd_for(255, 77, 77, "1")
        rq_wait_pos_spe_for_request(255, 77, 77, "1")
        rq_go_to("1")
        rq_wait("1")
        # end: URCap Program Node
        $ 1937 "Spatula_above" "noBreak"
        movel(Spatula_above_p, a=0.6, v=0.15)
        $ 1938 "Popup: Connect the vibration motor" "noBreak"
        popup("Connect the vibration motor", "Message", False, False, blocking=True)
        $ 1939 "tare_scale()" "noBreak"
        tare_scale()
        $ 1940 "container_start" "noBreak"
        movel(container_start_p, a=0.3, v=0.1)
        $ 1941 "container_wp_1" "noBreak"
        movel(container_wp_1_p, a=0.3, v=0.05)
        $ 1942 "Loop 1 times" "noBreak"
        Loop_9 = 0
        while (Loop_9 < 1):
          $ 1943 "Waypoint_55" "noBreak"
          global move_thread_flag_1943=0
          thread move_thread_1943():
            enter_critical
            move_thread_flag_1943 = 1
            movel(Waypoint_55_p, a=0.5, v=0.07)
            move_thread_flag_1943 = 2
            exit_critical
          end
          move_thread_flag_1943 = 0
          move_thread_han_1943 = run move_thread_1943()
          while (True):
            sleep(1.0E-10)
            if (move_thread_flag_1943 > 1):
              join move_thread_han_1943
              break
            end
            sync()
          end
          $ 1945 "Waypoint_56" "noBreak"
          movel(Waypoint_56_p, a=0.3, v=0.05)
          $ 1946 "Waypoint_74" "noBreak"
          movel(Waypoint_74_p, a=0.6, v=0.15)
          $ 1947 "Set AO[0]=3.0" "noBreak"
          set_standard_analog_out(0, 0.3)
          $ 1948 "Wait: 2.0" "noBreak"
          sleep(2.0)
          $ 1949 "Set AO[0]=0.0" "noBreak"
          set_standard_analog_out(0, 0.0)
          Loop_9 = Loop_9 + 1
        end
        $ 1953 "ftr_scoop2" "noBreak"
        movel(ftr_scoop2_p, a=0.3, v=0.05)
        $ 1954 "aftr_scoo3" "noBreak"
        movel(aftr_scoo3_p, a=0.3, v=0.05)
        $ 1955 "MoveJ" "noBreak"
        $ 1956 "Waypoint_60" "noBreak"
        movej(get_inverse_kin(Waypoint_60_p, qnear=Waypoint_60_q), a=0.5235987755982988, v=0.3490658503988659, r=0.05)
        $ 1957 "Waypoint_61" "noBreak"
        movej(get_inverse_kin(Waypoint_61_p, qnear=Waypoint_61_q), a=0.5235987755982988, v=0.3490658503988659, r=0.05)
        # begin: URCap Program Node
        #   Source: SensoPart VISOR Robotic, 2.0.0, SensoPart Industriesensorik GmbH
        #   Type: Approach Pose
        $ 1958 "Approach Pose" "noBreak"
        movej(pose_trans(easyPickPose,p[0.0000,0.0000,0.0500,0.0000,0.0000,0.0000]),a=0.4363,v=0.3491,t=0.000000,r=0.000000)
        # end: URCap Program Node
        # begin: URCap Program Node
        #   Source: SensoPart VISOR Robotic, 2.0.0, SensoPart Industriesensorik GmbH
        #   Type: Target Pose
        $ 1959 "Target Pose" "noBreak"
        movel(pose_trans(easyPickPose,p[0.0000,0.0000,-0.0000,0.0000,0.0000,0.0000]),a=0.1000,v=0.0500,t=0.000000,r=0.000000)
        # end: URCap Program Node
        $ 1960 "Close Gripper" "noBreak"
        $ 1961 "dispense_pos≔get_actual_tcp_pose()" "noBreak"
        global dispense_pos= get_actual_tcp_pose ()
        $ 1962 "MoveL" "noBreak"
        $ 1963 "Start_thread≔ True " "noBreak"
        global Start_thread=  True
        $ 1964 "vib_mot_thread≔ True " "noBreak"
        global vib_mot_thread=  True
        $ 1965 "tilt_angle≔current_pose[4]" "noBreak"
        global tilt_angle=current_pose[4]
        $ 1966 "Wait: 0.5" "noBreak"
        sleep(0.5)
        $ 1967 "Loop Weight_value≤Target_weight and tilt_angle≤-0.40" "noBreak"
        thread Thread_while_1967():
          while (True):
            $ 1968 "current_error≔Target_weight-Weight_value" "noBreak"
            global current_error=Target_weight-Weight_value
            $ 1969 "Integral_error≔Integral_error+current_error*dt" "noBreak"
            global Integral_error=Integral_error+current_error*dt
            $ 1970 "derivative≔(current_error-previous_error)/dt" "noBreak"
            global derivative=(current_error-previous_error)/dt
            $ 1971 "tilt_increment≔(kp*current_error)+(ki*Integral_error)+(kd*derivative)" "noBreak"
            global tilt_increment=(kp*current_error)+(ki*Integral_error)+(kd*derivative)
            $ 1972 "current_pose≔get_actual_tcp_pose()" "noBreak"
            global current_pose= get_actual_tcp_pose ()
            $ 1973 "tilt_angle≔current_pose[4]" "noBreak"
            global tilt_angle=current_pose[4]
            $ 1974 "tilt_pose≔pose_trans(current_pose, p[(tilt_increment/7), 0, 0, 0, tilt_increment, 0])" "noBreak"
            global tilt_pose=pose_trans(current_pose, p[(tilt_increment/7), 0, 0, 0, tilt_increment, 0])
            $ 1975 "movel(tilt_pose, a=0.025, v=0.015, r=0.00001)" "noBreak"
            movel(tilt_pose, a=0.025, v=0.015, r=0.00001)
            $ 1976 "previous_error≔current_error" "noBreak"
            global previous_error=current_error
          end
        end
        if (Weight_value <= Target_weight  and  tilt_angle <= -0.40):
          global thread_handler_1967=run Thread_while_1967()
          while (Weight_value <= Target_weight  and  tilt_angle <= -0.40):
            sync()
          end
          kill thread_handler_1967
        end
        $ 1977 "Start_thread≔ False " "noBreak"
        global Start_thread=  False
        $ 1979 "Weight_value≔get_weight()" "noBreak"
        global Weight_value=get_weight()
        $ 1980 "tilt_angle≔-1" "noBreak"
        global tilt_angle=-1
        $ 1981 "Wait: 0.5" "noBreak"
        sleep(0.5)
        $ 1982 "vib_mot_thread≔ False " "noBreak"
        global vib_mot_thread=  False
        $ 1983 "MoveL" "noBreak"
        $ 1984 "dispense_pos" "noBreak"
        movel(dispense_pos, a=0.2, v=0.05)
        $ 1985 "Integral_error≔0" "noBreak"
        global Integral_error=0
        $ 1986 "current_error≔0" "noBreak"
        global current_error=0
        $ 1987 "previous_error≔0" "noBreak"
        global previous_error=0
        $ 1988 "Set AO[0]=0.0" "noBreak"
        set_standard_analog_out(0, 0.0)
        # begin: URCap Program Node
        #   Source: SensoPart VISOR Robotic, 2.0.0, SensoPart Industriesensorik GmbH
        #   Type: Exit Pose
        $ 1989 "Exit Pose" "noBreak"
        movel(pose_trans(easyPickPose,p[0.0000,0.0000,-0.0000,0.0000,0.0000,0.0000]),a=0.5000,v=0.2500,t=0.000000,r=0.000000)
        # end: URCap Program Node
        easyPickObjTaken = True
      end
      # end: URCap Program Node
      # begin: URCap Program Node
      #   Source: SensoPart VISOR Robotic, 2.0.0, SensoPart Industriesensorik GmbH
      #   Type: No Object Detected
      $ 1990 "No Object Detected" "noBreak"
      if (visor_partsFound(easyPickVisorId) < 1):
        $ 1991 "Popup: No weigh scale detected" "noBreak"
        popup("No weigh scale detected", "Message", False, False, blocking=True)
        else:
      end
      # end: URCap Program Node
    end
    easyPickCount_4 = easyPickCount_4 + 1
    visor_easyPickUpdate(easyPickVisorId, "counter", easyPickCount_4)
    visor_easyPickSetIdent("a3cf6b", easyPickVisorId)
    # end: URCap Program Node
  end
  visorFuncEasyPick_5fe5fa()
  # end: URCap Program Node
  $ 1992 "powder dispensing"
  $ 1994 "Loop Weight_value<Target_weight"
  while (Weight_value<Target_weight):
    $ 1995 "MoveL"
    $ 1996 "Waypoint_75" "breakAfter"
    movel(Waypoint_75_p, a=0.3, v=0.05, r=0.05)
    $ 1997 "ftr_scoop2" "breakAfter"
    movel(ftr_scoop2_p, a=0.3, v=0.05)
    $ 1998 "aftr_scoop1" "breakAfter"
    movel(aftr_scoop1_p, a=0.3, v=0.05)
    $ 1999 "After_disp_3" "breakAfter"
    movel(After_disp_3_p, a=0.3, v=0.05)
    $ 2000 "Loop 1 times"
    Loop_13 = 0
    while (Loop_13 < 1):
      $ 2001 "Waypoint_55" "breakAfter"
      global move_thread_flag_2001=0
      thread move_thread_2001():
        enter_critical
        move_thread_flag_2001 = 1
        movel(Waypoint_55_p, a=0.5, v=0.07)
        move_thread_flag_2001 = 2
        exit_critical
      end
      move_thread_flag_2001 = 0
      move_thread_han_2001 = run move_thread_2001()
      while (True):
        sleep(1.0E-10)
        if (move_thread_flag_2001 > 1):
          join move_thread_han_2001
          break
        end
        sync()
      end
      $ 2003 "Waypoint_56" "breakAfter"
      movel(Waypoint_56_p, a=0.3, v=0.05)
      $ 2004 "Waypoint_74" "breakAfter"
      movel(Waypoint_74_p, a=0.3, v=0.05)
      $ 2005 "Set AO[0]=3.0"
      set_standard_analog_out(0, 0.3)
      $ 2006 "Wait: 2.0"
      sleep(2.0)
      $ 2007 "Set AO[0]=0.0"
      set_standard_analog_out(0, 0.0)
      Loop_13 = Loop_13 + 1
    end
    $ 2008 "ftr_scoop2" "breakAfter"
    movel(ftr_scoop2_p, a=0.3, v=0.05)
    $ 2009 "aftr_scoo3" "breakAfter"
    movel(aftr_scoo3_p, a=0.3, v=0.05)
    $ 2010 "MoveJ"
    $ 2011 "Waypoint_60" "breakAfter"
    movej(get_inverse_kin(Waypoint_60_p, qnear=Waypoint_60_q), a=0.5235987755982988, v=0.3490658503988659, r=0.05)
    $ 2012 "Waypoint_61" "breakAfter"
    movej(get_inverse_kin(Waypoint_61_p, qnear=Waypoint_61_q), a=0.5235987755982988, v=0.3490658503988659, r=0.05)
    $ 2013 "Waypoint_62" "breakAfter"
    movej(get_inverse_kin(Waypoint_62_p, qnear=Waypoint_62_q), a=0.5235987755982988, v=0.3490658503988659)
    $ 2014 "MoveL"
    $ 2015 "Start_thread≔ True "
    global Start_thread=  True
    $ 2016 "dispense_pos" "breakAfter"
    movel(dispense_pos, a=0.2, v=0.05)
    $ 2017 "vib_mot_thread≔ True "
    global vib_mot_thread=  True
    $ 2018 "Wait: 0.5"
    sleep(0.5)
    $ 2019 "Loop Weight_value≤Target_weight and tilt_angle≤-0.40"
    thread Thread_while_2019():
      while (True):
        $ 2020 "current_error≔Target_weight-Weight_value"
        global current_error=Target_weight-Weight_value
        $ 2021 "Integral_error≔Integral_error+current_error*dt"
        global Integral_error=Integral_error+current_error*dt
        $ 2022 "derivative≔(current_error-previous_error)/dt"
        global derivative=(current_error-previous_error)/dt
        $ 2023 "tilt_increment≔(kp*current_error)+(ki*Integral_error)+(kd*derivative)"
        global tilt_increment=(kp*current_error)+(ki*Integral_error)+(kd*derivative)
        $ 2024 "current_pose≔get_actual_tcp_pose()"
        global current_pose= get_actual_tcp_pose ()
        $ 2025 "tilt_angle≔current_pose[4]"
        global tilt_angle=current_pose[4]
        $ 2026 "tilt_pose≔pose_trans(current_pose, p[(tilt_increment/7), 0, 0, 0, tilt_increment, 0])"
        global tilt_pose=pose_trans(current_pose, p[(tilt_increment/7), 0, 0, 0, tilt_increment, 0])
        $ 2027 "movel(tilt_pose, a=0.025, v=0.015, r=0.00001)"
        movel(tilt_pose, a=0.025, v=0.015, r=0.00001)
        $ 2028 "previous_error≔current_error"
        global previous_error=current_error
        $ 2029 "Wait: 0.01"
        sleep(0.01)
      end
    end
    if (Weight_value <= Target_weight  and  tilt_angle <= -0.40):
      global thread_handler_2019=run Thread_while_2019()
      while (Weight_value <= Target_weight  and  tilt_angle <= -0.40):
        sync()
      end
      kill thread_handler_2019
    end
    $ 2030 "Start_thread≔ False "
    global Start_thread=  False
    $ 2031 "Set AO[0]=0.0"
    set_standard_analog_out(0, 0.0)
    $ 2032 "vib_mot_thread≔ False "
    global vib_mot_thread=  False
    $ 2034 "Weight_value≔get_weight()"
    global Weight_value=get_weight()
    $ 2035 "tilt_angle≔-1"
    global tilt_angle=-1
    $ 2036 "Wait: 0.5"
    sleep(0.5)
    $ 2037 "MoveL"
    $ 2038 "dispense_pos" "breakAfter"
    movel(dispense_pos, a=0.2, v=0.05)
    $ 2039 "Integral_error≔0"
    global Integral_error=0
    $ 2040 "current_error≔0"
    global current_error=0
    $ 2041 "previous_error≔0"
    global previous_error=0
  end
  $ 2042 "MoveL"
  $ 2043 "aftr_scoo3" "breakAfter"
  movel(aftr_scoo3_p, a=0.3, v=0.1)
  $ 2044 "ftr_scoop2" "breakAfter"
  movel(ftr_scoop2_p, a=0.4, v=0.1)
  $ 2045 "aftr_scoop1" "breakAfter"
  movel(aftr_scoop1_p, a=0.4, v=0.1)
  $ 2046 "After_disp_3" "breakAfter"
  movel(After_disp_3_p, a=0.4, v=0.1)
  $ 2047 "Set AO[0]=3.0"
  set_standard_analog_out(0, 0.3)
  $ 2048 "Wait: 2.0"
  sleep(2.0)
  $ 2049 "Set AO[0]=0.0"
  set_standard_analog_out(0, 0.0)
  $ 2050 "aftr_scoop1" "breakAfter"
  movel(aftr_scoop1_p, a=1.2, v=0.25)
  $ 2051 "ftr_scoop2" "breakAfter"
  movel(ftr_scoop2_p, a=0.4, v=0.1)
  $ 2052 "Waypoint_63" "breakAfter"
  movel(Waypoint_63_p, a=1.2, v=0.25, r=0.05)
  $ 2053 "Start" "breakAfter"
  movel(Start_p, a=0.6, v=0.15)
  $ 2054 "Popup: Powder dispensed successfully..."
  popup("Powder dispensed successfully...", "Message", False, False, blocking=True)
  elif (38 == switch_1):
    $ 2055 "Case 38"
    $ 2056 "PowderA(M200)"
    # begin: URCap Program Node
    #   Source: SensoPart VISOR Robotic, 2.0.0, SensoPart Industriesensorik GmbH
    #   Type: VISOR Robotic App
    $ 2057 "VISOR Easy Pick"
    def visorFuncEasyPick_5cb6a0():
      # begin: URCap Program Node
      #   Source: SensoPart VISOR Robotic, 2.0.0, SensoPart Industriesensorik GmbH
      #   Type: Easy Pick Setup
      $ 2058 "# 1 Setup" "noBreak"
      local easyPickVisorId = 1
      local easyPickArmMounted = True
      local easyPickSetJob = True
      local easyPickJobName = "PowderA"
      local easyPickAtImgAcq = False
      local easyPickImgAcqPose = cont_img_pose
      # end: URCap Program Node
      # begin: URCap Program Node
      #   Source: SensoPart VISOR Robotic, 2.0.0, SensoPart Industriesensorik GmbH
      #   Type: Process
      $ 2059 "Process" "noBreak"
      local easyPickObjTaken = False
      local easyPickTrigger = False
      local easyPickPoseIdx = 0
      local easyPickPose = p[0,0,0,0,0,0]
      def easyPickFuncTrigger(visorId, setJob, jobName, arm):
      if (setJob):
        visor_changeJob(visorId, jobName, 6000)
      end
      if (arm):
        visor_trigger(visorId, 6000, "arm")
      else:
        visor_trigger(visorId, 6000)
      end
      global easyPickParts_6=visor_partsFound(visorId)
      visor_easyPickUpdate(visorId, "parts", visor_partsFound(visorId))
      return visor_getPose3d(visorId, 0)
    end
    while (not easyPickObjTaken):
      easyPickTrigger = (easyPickCount_6 >= visor_partsFound(easyPickVisorId)) or (easyPickCount_6 > 9) or (not visor_easyPickCheckIdent("38655b", easyPickVisorId))
      if (easyPickTrigger):
        easyPickCount_6 = 0
      end
      easyPickPoseIdx = easyPickCount_6
      easyPickPose = visor_getPose3d(easyPickVisorId, easyPickPoseIdx)
      visor_easyPickUpdate(easyPickVisorId, "counter", easyPickPoseIdx)
      # begin: URCap Program Node
      #   Source: SensoPart VISOR Robotic, 2.0.0, SensoPart Industriesensorik GmbH
      #   Type: Image Acquisition Pose
      $ 2060 "Image Acquisition Pose" "noBreak"
      if (easyPickTrigger):
        if (not easyPickAtImgAcq):
          movej(pose_trans(easyPickImgAcqPose,p[0.0000,0.0000,-0.0000,0.0000,0.0000,0.0000]),a=1.3963,v=1.0472,t=0.000000,r=0.000000)
          easyPickAtImgAcq = True
        end
        easyPickPose = easyPickFuncTrigger(easyPickVisorId, easyPickSetJob, easyPickJobName, easyPickArmMounted)
      end
      # end: URCap Program Node
      # begin: URCap Program Node
      #   Source: SensoPart VISOR Robotic, 2.0.0, SensoPart Industriesensorik GmbH
      #   Type: Object Detected
      $ 2061 "Object Detected" "noBreak"
      if (visor_partsFound(easyPickVisorId) > 0):
        $ 2062 "Open Gripper" "noBreak"
        # begin: URCap Program Node
        #   Source: Robotiq_Grippers, 1.8.4.4844, Robotiq Inc.
        #   Type: Gripper
        $ 2063 "Gripper Open (1)" "noBreak"
        if not(gripper_connected[0]):
          popup("Gripper 1 must be connected to run this program.", "No connection", False, True, True)
        end
        if not(rq_is_gripper_activated("1")):
          popup("Gripper 1 is not activated. Go to Installation tab > Gripper to activate it and run the program again.", "Not activated", False, True, True)
        end
        rq_set_pos_spd_for(0, 77, 77, "1")
        rq_wait_pos_spe_for_request(0, 77, 77, "1")
        rq_go_to("1")
        rq_wait("1")
        # end: URCap Program Node
        $ 2064 "MoveJ" "noBreak"
        $ 2065 "Waypoint_76" "noBreak"
        movej(get_inverse_kin(Waypoint_76_p, qnear=Waypoint_76_q), a=1.3962634015954636, v=1.0471975511965976)
        # begin: URCap Program Node
        #   Source: SensoPart VISOR Robotic, 2.0.0, SensoPart Industriesensorik GmbH
        #   Type: Approach Pose
        $ 2066 "Approach Pose" "noBreak"
        movej(pose_trans(easyPickPose,p[0.0000,0.0000,0.0500,0.0000,0.0000,0.0000]),a=1.3963,v=1.0472,t=0.000000,r=0.000000)
        # end: URCap Program Node
        # begin: URCap Program Node
        #   Source: SensoPart VISOR Robotic, 2.0.0, SensoPart Industriesensorik GmbH
        #   Type: Target Pose
        $ 2067 "Target Pose" "noBreak"
        movel(pose_trans(easyPickPose,p[0.0000,0.0000,-0.0000,0.0000,0.0000,0.0000]),a=0.5000,v=0.2500,t=0.000000,r=0.000000)
        # end: URCap Program Node
        $ 2068 "Close Gripper" "noBreak"
        # begin: URCap Program Node
        #   Source: Robotiq_Grippers, 1.8.4.4844, Robotiq Inc.
        #   Type: Gripper
        $ 2069 "Gripper Move0mm (1)" "noBreak"
        if not(gripper_connected[0]):
          popup("Gripper 1 must be connected to run this program.", "No connection", False, True, True)
        end
        if not(rq_is_gripper_activated("1")):
          popup("Gripper 1 is not activated. Go to Installation tab > Gripper to activate it and run the program again.", "Not activated", False, True, True)
        end
        rq_set_pos_spd_for(247, 77, 77, "1")
        rq_wait_pos_spe_for_request(247, 77, 77, "1")
        rq_go_to("1")
        rq_wait("1")
        # end: URCap Program Node
        # begin: URCap Program Node
        #   Source: SensoPart VISOR Robotic, 2.0.0, SensoPart Industriesensorik GmbH
        #   Type: Exit Pose
        $ 2070 "Exit Pose" "noBreak"
        movel(pose_trans(easyPickPose,p[0.0000,0.0000,0.0500,0.0000,0.0000,0.0000]),a=0.5000,v=0.2500,t=0.000000,r=0.000000)
        # end: URCap Program Node
        easyPickObjTaken = True
      end
      # end: URCap Program Node
      # begin: URCap Program Node
      #   Source: SensoPart VISOR Robotic, 2.0.0, SensoPart Industriesensorik GmbH
      #   Type: No Object Detected
      $ 2071 "No Object Detected" "noBreak"
      if (visor_partsFound(easyPickVisorId) < 1):
        $ 2072 "Popup: No Powder container is detected" "noBreak"
        popup("No Powder container is detected", "Message", False, False, blocking=True)
        else:
      end
      # end: URCap Program Node
    end
    easyPickCount_6 = easyPickCount_6 + 1
    visor_easyPickUpdate(easyPickVisorId, "counter", easyPickCount_6)
    visor_easyPickSetIdent("38655b", easyPickVisorId)
    # end: URCap Program Node
  end
  visorFuncEasyPick_5cb6a0()
  # end: URCap Program Node
  $ 2073 "MoveJ"
  $ 2074 "PowderA_wayp1" "breakAfter"
  movej(get_inverse_kin(PowderA_wayp1_p, qnear=PowderA_wayp1_q), a=1.3962634015954636, v=1.0471975511965976, r=0.05)
  $ 2075 "MoveL"
  $ 2076 "Waypoint_80" "breakAfter"
  movel(Waypoint_80_p, a=1.2, v=0.25)
  $ 2077 "MoveL"
  $ 2078 "Decapp_above" "breakAfter"
  movel(Decapp_above_p, a=1.2, v=0.25)
  $ 2079 "Set GRP_3F_Open=On"
  set_standard_digital_out(5, True)
  $ 2080 "Wait: 0.5"
  sleep(0.5)
  $ 2081 "Decapp_place" "breakAfter"
  movel(Decapp_place_p, a=0.3, v=0.05)
  $ 2082 "Set GRP_3F_Open=Off"
  set_standard_digital_out(5, False)
  $ 2083 "Wait: 0.5"
  sleep(0.5)
  # begin: URCap Program Node
  #   Source: Robotiq_Grippers, 1.8.4.4844, Robotiq Inc.
  #   Type: Gripper
  $ 2084 "Gripper Move40mm (1)"
  if not(gripper_connected[0]):
    popup("Gripper 1 must be connected to run this program.", "No connection", False, True, True)
  end
  if not(rq_is_gripper_activated("1")):
    popup("Gripper 1 is not activated. Go to Installation tab > Gripper to activate it and run the program again.", "Not activated", False, True, True)
  end
  rq_set_pos_spd_for(64, 77, 77, "1")
  rq_wait_pos_spe_for_request(64, 77, 77, "1")
  rq_go_to("1")
  rq_wait("1")
  # end: URCap Program Node
  $ 2085 "MoveL"
  $ 2086 "Decapp_above" "breakAfter"
  movel(Decapp_above_p, a=1.2, v=0.25)
  $ 2087 "Waypoint_78" "breakAfter"
  movel(Waypoint_78_p, a=1.2, v=0.25, r=0.05)
  $ 2088 "Home (Safe)"
  movej([-1.2302089344500047, -1.2969853503591224, -1.875639182904262, -1.539621866126728, 1.5731943360401213, -2.80099559440227], a=1.3962634015954636, v=1.0471975511965976)
  elif (39 == switch_1):
    $ 2089 "Case 39"
    $ 2090 "Decap Container A"
    $ 2091 "MoveL"
    $ 2092 "Waypoint_81" "breakAfter"
    movel(Waypoint_81_p, a=1.2, v=0.25)
    $ 2093 "Waypoint_79" "breakAfter"
    movel(Waypoint_79_p, a=1.2, v=0.25)
    # begin: URCap Program Node
